// iterate untill diff < epsilon or i_max=7 is reached
// 5 passes converge to <0.25" for the normal operating envelope (alt >= 3deg);
// see testing/check_pointing_inversion.py. Kept a small margin over the bare minimum.
bValid := FALSE;
FOR i:=0 TO 7 BY 1 DO
	d_ha := d_ha_new;
	d_dec := d_dec_new;
	fbpointing(
		HourAngle := LMOD(HourAngle-d_ha,360),
		Declination:= Declination-d_dec,
		Latitude:= Latitude,
		HourAngle_correction => d_ha_new,
		Declination_correction => d_dec_new
	);
	IF ABS(d_ha - d_ha_new) <= epsilon/3600.0 AND ABS(d_dec - d_dec_new) <= epsilon/3600.0 THEN
		bValid := TRUE;
		EXIT;
	END_IF
END_FOR;
// below alt~2-3deg the map is chaotic and never settles within epsilon (see script above);
// do not hand back whatever the last unconverged pass produced
IF bValid THEN
	HourAngle_correction := d_ha_new;
	Declination_correction := d_dec_new;
ELSE
	HourAngle_correction := 0.0;
	Declination_correction := 0.0;
END_IF

END_FUNCTION_BLOCK

// ---- POUs/FB_HomeDropReason.TcPOU
// Why a pending home was dropped after 2 min (#108): the text for the home end state and the WARN. Pure logic,
// tested offline in IAG50cmTests (#120). Order matters: not ready wins over a stop that did not finish.
FUNCTION_BLOCK FB_HomeDropReason
VAR_INPUT
	bReady			: BOOL;		// telescope ready
	bStopPending	: BOOL;		// TCS_command is stop, or the telescope is not at rest
END_VAR
VAR_OUTPUT
	sEnd			: STRING(40);
	sWhy			: STRING(160);
END_VAR

IF NOT bReady THEN
	sEnd := 'cancelled: telescope not ready';
	sWhy := 'the telescope was not ready for 2 min. Power on, then send the home again.';
ELSIF bStopPending THEN
	sEnd := 'cancelled: stop did not finish';
	sWhy := 'the stop before the home did not finish within 2 min. Send the stop, then the home again.';
ELSE
	sEnd := 'cancelled: axes busy';
	sWhy := 'the axes were busy for 2 min. Send the home again.';
END_IF

END_FUNCTION_BLOCK

// ---- POUs/FB_SweepStop.TcPOU
// A stop in the calibration sweep (#113): the axes stay enabled and uncalibrated, the sweep is aborted by the stop. Once the
// stop has settled (for 3 scans) and no homing is running any more, the uncalibrated axes are switched off for one scan, so
// the telescope ends like a stop in the covers phase (READY_STATE -2, no error) and the next power-on starts the sweep
// again. Calibrated axes stay enabled. Pure logic, tested offline in IAG50cmTests.
// #197: ArmAll() is the same for a park without a completed power-on (the axes are on, but the telescope can never be
// ready): every axis is switched off once at rest, calibrated or not, and the axes-off park then parks in place.
FUNCTION_BLOCK FB_SweepStop
VAR_INPUT
	bSettled		: BOOL;		// FB_TelescopeControl.bSettled: at rest and no stop transaction running
	bHaCalibrated	: BOOL;
	bDecCalibrated	: BOOL;
	bHaHoming		: BOOL;		// FB_LatchHome.Busy
	bDecHoming		: BOOL;
	bOtherBusy		: BOOL;		// #197: the focus is moving; waited for in the all-axes mode only
END_VAR
VAR_OUTPUT
	bDisableHa		: BOOL;		// one scan
	bDisableDec		: BOOL;
END_VAR
VAR
	bPending		: BOOL;
	bAll			: BOOL;		// #197: switch every axis off, not only the uncalibrated ones
	nSettledScans	: UINT;
END_VAR
VAR CONSTANT
	nConfirmScans	: UINT := 3;
END_VAR

bDisableHa := FALSE;
bDisableDec := FALSE;
IF bPending THEN
	IF bSettled AND NOT bHaHoming AND NOT bDecHoming AND NOT (bAll AND bOtherBusy) THEN
		IF nSettledScans < nConfirmScans THEN
			nSettledScans := nSettledScans + 1;
		END_IF
	ELSE
		nSettledScans := 0;
	END_IF
	IF nSettledScans >= nConfirmScans THEN
		bDisableHa := bAll OR NOT bHaCalibrated;
		bDisableDec := bAll OR NOT bDecCalibrated;
		bPending := FALSE;
		bAll := FALSE;
	END_IF
END_IF

// A stop arrived in the calibration sweep (power-on stage 40 or later).
METHOD Arm
IF NOT (bPending AND bAll) THEN	// a pending ArmAll() is not narrowed
	bPending := TRUE;
	nSettledScans := 0;
END_IF
END_METHOD

// A park without a completed power-on (#197): switch every axis off once at rest. Idempotent: it may be called every scan.
METHOD ArmAll
IF NOT (bPending AND bAll) THEN
	bPending := TRUE;
	bAll := TRUE;
	nSettledScans := 0;
END_IF
END_METHOD

// Error, reset or a new power-on: nothing to switch off any more.
METHOD Cancel
bPending := FALSE;
bAll := FALSE;
nSettledScans := 0;
END_METHOD

END_FUNCTION_BLOCK

// ---- POUs/Functions/F_HourAngleOffsetOnAxis.TcPOU
// Hour-angle-axis correction (degrees) for a cross-declination offset on the sky (fHourAngleOffset, degrees) at
// declination fDeclination (degrees): fHourAngleOffset / COS(fDeclination). Near the pole 1/COS grows without bound
// and is a division by zero at +-90 deg, so COS is floored at COS(89.5 deg) (factor 115 at most) and the result is
// limited to +-10 deg, the bound BROTLib puts on the offset command (BROTLib#27, same as MONETcommon's
// F_AzimuthOffsetOnAxis near the zenith). Below |dec| = 89.5 deg the result is unchanged.
FUNCTION F_HourAngleOffsetOnAxis : LREAL
VAR_INPUT
	fHourAngleOffset	: LREAL;	// cross-declination offset on the sky, degrees
	fDeclination		: LREAL;	// declination, degrees
END_VAR
VAR CONSTANT
	D2R				: LREAL := 0.017453292519943295;
	MIN_COS			: LREAL := 0.008726535498373935;	// COS(89.5 deg)
	MAX_AXIS_OFFSET	: LREAL := 10.0;					// degrees
END_VAR

F_HourAngleOffsetOnAxis := LIMIT(-MAX_AXIS_OFFSET, fHourAngleOffset / MAX(COS(fDeclination * D2R), MIN_COS), MAX_AXIS_OFFSET);

END_FUNCTION

// ---- POUs/DomeControl/FB_DomeControl.TcPOU
FUNCTION_BLOCK FB_DomeControl IMPLEMENTS I_Dome
VAR_INPUT
	ipTelescope: I_RaDecTelescope;
END_VAR
VAR
	ipState		: I_DomeState := fbDomeIdleState;
	bOpen		: BOOL;
	bClose		: BOOL;
	bReset		: BOOL;
	bHome		: BOOL;
	bTrack		: BOOL;
	bPark		: BOOL;
	bStop		: BOOL;
	bStopDone	: BOOL;
	
	fDomeAziGoInput			: LREAL := 180.0;
	fDomeAziGo				: LREAL := 180.0;
	fDomeAziCurrent			: LREAL := 0.0;
	eDomeRotationState		: E_DomeRotationState;
	eDomeRotationStateOld	: E_DomeRotationState;
	eDomeShutterState		: E_RoofState;
	eDomeShutterStateOld	: E_RoofState;
	bParked			: BOOL;
	
	bDomeError	: BOOL;
	iDomeErrorID: UINT;
	
	ipStateOld			: I_DomeState := fbDomeIdleState;
	fbDomeCloseingState : FB_DomeClosingState(THIS);
	fbDomeErrorState	: FB_DomeErrorState(THIS);
	fbDomeHomeingState	: FB_DomeHomingState(THIS);
	fbDomeIdleState		: FB_DomeIdleState(THIS);
	fbDomeOpeningState	: FB_DomeOpeningState(THIS);
	fbDomeMovingState	: FB_DomeMovingState(THIS);
	fbDomeParkingState	: FB_DomeParkingState(THIS);
	fbDomeStoppingState	: FB_DomeStoppingState(THIS);
	

	rtrigOpen		: R_TRIG;
	rtrigClose		: R_TRIG;
	rtrigReset		: R_TRIG;
	rtrigHome		: R_TRIG;
	rtrigPark		: R_TRIG;
	rtrigStop		: R_TRIG;
	
	fbComm			: I_Comm;
	tonComm 		: TON := (PT:=T#5S);
	
	fbDomeParkedEvent:	FB_EventLog;
	fbDomeStopEvent:	FB_EventLog;
	fbDomeErrorEvent: FB_EventLog;
	
	sSendstring	: STRING;
	Stage		: UINT:= 0;
	Timer		: TON := (PT:=T#30S);
	fbSend		: SendString;
	bSendBusy	: BOOL;
	eSendErrorID: ComError_t;

	fbReceive		: ReceiveString;
	sReceivedString	: STRING;
	sLastReceivedString: STRING;
	bStringReceived	: BOOL;
	bReceiveBusy	: BOOL;
	bReceiveError	: BOOL;
	eReceiveErrorID	: ComError_t;
	bReceiveTimeout	: BOOL;
END_VAR
VAR CONSTANT
	nCapabilities : INT := 2; 	//OPEN TSI : TELESCOPE.CONFIG.CAPABILITIES
END_VAR

// account for off center mount
IF fDomeAziGoInput >= 0.0 AND fDomeAziGoInput < 115.0 THEN
	fDomeAziGo := fDomeAziGoInput - 5.0;
ELSIF fDomeAziGoInput >= 225.0 AND fDomeAziGoInput < 360.0 THEN
	fDomeAziGo := fDomeAziGoInput + 5.0;
ELSE
	fDomeAziGo := fDomeAziGoInput;
END_IF

//	Receive string data:
fbReceive(
	Prefix:='',
	Suffix:= '',
	Timeout:= T#1S,
	ReceivedString:= sReceivedString,
	RXbuffer:= RxBufferDome,
	StringReceived=> bStringReceived,
	Busy=> bReceiveBusy,
	Error=> ,
	RxTimeout=> bReceiveTimeout );
// Check Errors
IF fbSend.Error <> COMERROR_NOERROR THEN
	eSendErrorID := fbSend.Error;
	bDomeError := TRUE;
END_IF
IF fbReceive.Error <> COMERROR_NOERROR THEN
	eReceiveErrorID := fbReceive.Error;
	bDomeError := TRUE;
END_IF

IF bDomeError THEN
	THIS^.ipState.FoundError();
END_IF

rtrigOpen(CLK := bOpen);
rtrigClose(CLK := bClose);
rtrigReset(CLK := bReset);
rtrigHome(CLK := bHome);
rtrigPark(CLK := bPark);
rtrigStop(CLK := bStop);

// #96: a stop wins over every other request of the same scan, which are dropped with it
IF (rtrigStop.Q) THEN
	bStop := FALSE;
	bOpen := FALSE;
	bClose := FALSE;
	bHome := FALSE;
	bPark := FALSE;
	bTrack := FALSE;
	ipState.StopCommand();
END_IF

IF (rtrigReset.Q) THEN
	bReset := FALSE;
	ipState.ResetCommand();
END_IF

IF (rtrigClose.Q) THEN
	bClose := FALSE;
	ipState.CloseCommand();
END_IF

IF (rtrigOpen.Q) THEN
	bOpen := FALSE;
	ipState.OpenCommand();
END_IF

IF (rtrigHome.Q) THEN
	bHome := FALSE;
	ipState.HomeCommand();
END_IF

IF (rtrigPark.Q) THEN
	bPark := FALSE;
	bTrack := FALSE;
	ipState.ParkCommand();
END_IF

// #83: requests are one-shot, like the covers (#66). They are consumed in this scan whether they produced an edge or
// not: a caller repeating a request every scan gave a single edge and then left the flag TRUE, so no later request of
// that kind had an edge until a PLC restart.
bOpen := FALSE;
bClose := FALSE;
bReset := FALSE;
bHome := FALSE;
bPark := FALSE;
bStop := FALSE;

bStopDone := FALSE;
ipState.RunState();

IF eDomeRotationState = E_DomeRotationState.parked AND eDomeShutterState = E_RoofState.closed THEN
	bParked := TRUE;
ELSE
	bParked := FALSE;
END_IF
// send telemetry
tonComm(IN:=TRUE);
IF tonComm.Q THEN // publish new payload every 5 seconds
	tonComm(IN:=FALSE);
	THIS^._SendTelemetry();	
END_IF


fbDomeParkedEvent(
	Trigger := bParked,
	Level := ADSLOG_MSGTYPE_HINT,
	OnMessage := 'Dome is in parking position and closed.',
	comm:= fbComm);
fbDomeStopEvent(
	Trigger := bStopDone,
	Level := ADSLOG_MSGTYPE_HINT,
	OnMessage := 'Dome stopped: rotation holds the current azimuth, a shutter movement is not stopped.',
	comm:= fbComm);
fbDomeErrorEvent(
	Trigger := bDomeError,
	Level := ADSLOG_MSGTYPE_ERROR,
	FormatString := 'Dome Error %s',
	OnMessage := 'found.',
	OffMessage := 'resolved.',
	comm:= fbComm);
// Buffer
ipStateOld := ipState;
eDomeRotationStateOld := eDomeRotationState;
eDomeShutterStateOld := eDomeShutterState;

PROPERTY _DomeRotationState : E_DomeRotationState
GET
_DomeRotationState := eDomeRotationState;
END_GET
SET
eDomeRotationState := _DomeRotationState;
END_SET
END_PROPERTY

PROPERTY _DomeShutterState : E_RoofState
GET
_DomeShutterState := eDomeShutterState;
END_GET
SET
eDomeShutterState := _DomeShutterState;
END_SET
END_PROPERTY

PROPERTY  _Error : BOOL
GET
_Error := bDomeError;
END_GET
SET
bDomeError := _Error;
END_SET
END_PROPERTY

PROPERTY _StopDone : BOOL
GET
_StopDone := bStopDone;
END_GET
SET
bStopDone := _StopDone;
END_SET
END_PROPERTY

PROPERTY _HasReceivedString : Bool
GET
_HasReceivedString := bStringReceived;
END_GET
SET
END_SET
END_PROPERTY

PROPERTY _Parked : BOOL
GET
_Parked := bParked;
END_GET
SET
bParked := _Parked;
END_SET
END_PROPERTY

PROPERTY _Position : LREAL
GET
_Position := fDomeAziGo;
END_GET
SET
fDomeAziCurrent := _Position;
END_SET
END_PROPERTY

PROPERTY _ReceivedString : STRING
GET
_ReceivedString := sReceivedString;
END_GET
SET
END_SET
END_PROPERTY

METHOD _SendTelemetry : BOOL
VAR_INPUT
END_VAR
IF eDomeShutterState = E_RoofState.opened THEN
	fbComm.PublishLREAL('telescope', 'dome', 'AUXILIARY.DOME.REALPOS', 1.0);
ELSIF eDomeShutterState = E_RoofState.closing OR eDomeShutterState = E_RoofState.opening OR eDomeShutterState = E_RoofState.unknown THEN
	fbComm.PublishLREAL('telescope', 'dome', 'AUXILIARY.DOME.REALPOS', 0.5);
ELSIF eDomeShutterState = E_RoofState.closed THEN
	fbComm.PublishLREAL('telescope', 'dome', 'AUXILIARY.DOME.REALPOS', 0.0);
ELSE
	fbComm.PublishLREAL('telescope', 'dome', 'AUXILIARY.DOME.REALPOS', -1.0);
END_IF

IF ipState.StateID = 'Opening State' THEN
	fbComm.PublishLREAL('telescope', 'dome', 'AUXILIARY.DOME.TARGETPOS', 1.0);
ELSE
	fbComm.PublishLREAL('telescope', 'dome', 'AUXILIARY.DOME.TARGETPOS', 0.0);
END_IF

IF bDomeError THEN
	fbComm.PublishINT('telescope', 'dome', 'AUXILIARY.DOME.ERROR_STATE', 1);
	fbComm.PublishLREAL('telescope', 'dome', 'AUXILIARY.DOME.READY_STATE', -1.0);
ELSE
	fbComm.PublishINT('telescope', 'dome', 'AUXILIARY.DOME.ERROR_STATE', 0);
	IF bParked THEN
		fbComm.PublishLREAL('telescope', 'dome', 'AUXILIARY.DOME.READY_STATE', 0.0);
	ELSIF bTrack THEN
		fbComm.PublishLREAL('telescope', 'dome', 'AUXILIARY.DOME.READY_STATE', 8.0);
	ELSE
		fbComm.PublishLREAL('telescope', 'dome', 'AUXILIARY.DOME.READY_STATE', 1.0);
	END_IF
END_IF

IF eDomeRotationState = E_DomeRotationState.slewing OR eDomeRotationState = E_DomeRotationState.unknown THEN
	fbComm.PublishLREAL('telescope', 'dome', 'AUXILIARY.DOME.MOTION_STATE', 1.0);
ELSE
	fbComm.PublishLREAL('telescope', 'dome', 'AUXILIARY.DOME.MOTION_STATE', 0.0);
END_IF
fbComm.PublishLREAL('telescope', 'dome', 'AUXILIARY.DOME.AZ', THIS^.Position);
END_METHOD

PROPERTY _Track : BOOL
GET
_Track := bTrack;
END_GET
END_PROPERTY

PROPERTY Capabilities : INT
GET
Capabilities := nCapabilities;
END_GET
END_PROPERTY

METHOD Close : BOOL
VAR_INPUT
END_VAR
bClose:=True;
END_METHOD

PROPERTY Closed : BOOL
GET
END_GET
END_PROPERTY

PROPERTY Error : Bool
GET
Error := bDomeError;
END_GET
END_PROPERTY

PROPERTY ErrorID : UDINT
GET
END_GET
END_PROPERTY

//FB_Init is always available implicitly and it is used primarily for initialization.
//The return value is not evaluated. For a specific influence, you can also declare the
//methods explicitly and provide additional code there with the standard initialization
//code. You can evaluate the return value.
METHOD FB_Init: BOOL
VAR_INPUT
    bInitRetains	: BOOL; // TRUE: the retain variables are initialized (reset warm / reset cold)
    bInCopyCode		: BOOL;  // TRUE: the instance will be copied to the copy code afterward (online change)
	comm			: I_Comm;
END_VAR
THIS^.fbComm 				:= comm;
END_METHOD

METHOD Open : BOOL
VAR_INPUT
END_VAR
bOpen := True;
END_METHOD

PROPERTY Opened : BOOL
GET
END_GET
END_PROPERTY

METHOD Park : BOOL
VAR_INPUT
END_VAR
bPark := TRUE;
END_METHOD

PROPERTY Parked : BOOL
GET
Parked := bParked;
END_GET
END_PROPERTY

PROPERTY Position : LREAL
GET
Position := fDomeAziCurrent;
END_GET
SET
fDomeAziGoInput := Position;
END_SET
END_PROPERTY

METHOD Reset : BOOL
VAR_INPUT
END_VAR
bReset := True;
END_METHOD

PROPERTY RotState : E_DomeRotationState
GET
RotState := eDomeRotationState;
END_GET
END_PROPERTY

METHOD SetState : BOOL
VAR_INPUT
	newState :I_DomeState;
END_VAR
THIS^.ipState := newState;
END_METHOD

{warning 'add property implementation'}
PROPERTY ShutterState : BROTLib.E_RoofState
GET
END_GET
SET
END_SET
END_PROPERTY

PROPERTY Slewing : BOOL
GET
END_GET
END_PROPERTY

METHOD Stop : BOOL
VAR_INPUT
END_VAR
// #96: the dome has no stop command, the state holds the azimuth it reads (FB_DomeStoppingState)
bStop := TRUE;
END_METHOD

METHOD StopTrack : BOOL
VAR_INPUT
END_VAR
bTrack := FALSE;
END_METHOD

METHOD Track : BOOL
VAR_INPUT
END_VAR
bTrack := TRUE;
END_METHOD

PROPERTY Tracking : BOOL
GET
Tracking := bTrack;
END_GET
END_PROPERTY

END_FUNCTION_BLOCK

// ---- POUs/DomeControl/States/FB_DomeClosingState.TcPOU
FUNCTION_BLOCK FB_DomeClosingState EXTENDS  FB_DomeState
VAR
	Stage		: UINT:= 0;
	tonSleep	: TON := (PT:=T#5S);
	tonTimeout	: TON:= (PT:=T#3M); // see Baader Handbook
	// #202: d#closhut is acknowledged (d#gotmess) but the shutter stays open (d#shutope): the command is sent again at
	// most nMaxAttempts times in all, then it is an error. Before, it was sent for ever, because the timeout is stopped
	// at every poll, and nothing was logged.
	nAttempts	: UINT;
	nMaxAttempts: UINT := 3;
END_VAR


METHOD CloseCommand : BOOL
// #202: a new close starts the shutter command again, with a fresh count
LogEvent(sText := 'Dome: close received while closing, the shutter command is started again', sLevel := 'WARNING');
nAttempts := 0;
Stage := 0;
tonSleep(IN:=FALSE);
tonTimeout(IN:=FALSE);
END_METHOD

METHOD FoundError : BOOL
nAttempts := 0;
Stage:= 0;
tonSleep(IN:=FALSE);
tonTimeout(IN:=FALSE);
pDome^._Error := TRUE;
pDome^.SetState(pDome^.fbDomeErrorState);
END_METHOD


METHOD OpenCommand : BOOL
nAttempts := 0;
Stage:= 0;
tonSleep(IN:=FALSE);
tonTimeout(IN:=FALSE);
pDome^.SetState(pDome^.fbDomeOpeningState);
END_METHOD

METHOD RunState : BOOL
VAR_INPUT
END_VAR
CASE Stage OF
	0:
		tonTimeout(IN:=TRUE);
		Stage := 1;
	1:
		pDome^.fbSend(	SendString:= 'd#closhut',
					TXbuffer:= TxBufferDome,
					Busy=>,
					Error=> );
		IF NOT pDome^.fbSend.Busy  THEN
			Stage := 2;
		END_IF
	2:
		IF pDome^.bStringReceived THEN
			IF pDome^._ReceivedString = 'd#comerro' OR pDome^._ReceivedString = 'd#domerro' THEN
				foundError();
			ELSIF pDome^._ReceivedString = 'd#gotmess' THEN
				Stage := 3;
			END_IF
		ELSIF NOT pDome^.fbReceive.Busy THEN
			tonSleep(IN:=TRUE);
			IF tonSleep.Q THEN
				tonSleep(IN:=FALSE);
				Stage := 1;
			END_IF
		END_IF
		tonTimeout(IN:=TRUE);
		IF tonTimeout.Q THEN
			tonTimeout(IN:=FALSE);
			foundError();
		END_IF
	3:
		tonTimeout(IN:=FALSE);
		
		tonSleep(IN:=TRUE);
		IF tonSleep.Q THEN
			tonSleep(IN:=FALSE);
			Stage := 4;
			tonTimeout(IN:=TRUE);
		END_IF
	4:
		pDome^.fbSend(	SendString:= 'd#getshut',
					TXbuffer:= TxBufferDome,
					Busy=>,
					Error=> );
		IF NOT pDome^.fbSend.Busy  THEN
			Stage := 5;
		END_IF
	5: 
		IF pDome^.bStringReceived THEN
			IF pDome^._ReceivedString = 'd#comerro' OR pDome^._ReceivedString = 'd#domerro' THEN
				FoundError();
			ELSIF pDome^._ReceivedString = 'd#shutclo' THEN
				pDome^._DomeShutterState := E_RoofState.closed;
				Stage := 6;
			ELSIF pDome^._ReceivedString = 'd#shutope' THEN
				pDome^._DomeShutterState := E_RoofState.opened;
				nAttempts := nAttempts + 1;
				IF nAttempts >= nMaxAttempts THEN
					LogEvent(sText := 'Dome: the shutter does not close, d#closhut is acknowledged but the shutter stays open', sLevel := 'WARNING');
					FoundError();
				ELSE
					Stage := 0;
				END_IF
			ELSIF pDome^._ReceivedString = 'd#shutrun' THEN
				pDome^._DomeShutterState := E_RoofState.closing;
				Stage := 3;
			END_IF
		ELSIF NOT pDome^.fbReceive.Busy THEN
			// mixed up string? ask again
			tonSleep(IN:=TRUE);
			IF tonSleep.Q THEN
				tonSleep(IN:=FALSE);
				Stage := 4;
			END_IF
		END_IF
		tonTimeout(IN:=TRUE);
		IF tonTimeout.Q THEN
			tonTimeout(IN:=FALSE);
			FoundError();
		END_IF
	
	6:
		tonTimeout(IN:=FALSE);
		SuccessfulFinished();
		
END_CASE
END_METHOD


PROPERTY StateID : STRING
GET
StateID := 'Closing State';
END_GET
END_PROPERTY


METHOD SuccessfulFinished : BOOL
nAttempts := 0;
Stage:= 0;
tonSleep(IN:=FALSE);
tonTimeout(IN:=FALSE);
pDome^.SetState(pDome^.fbDomeIdleState);
END_METHOD

END_FUNCTION_BLOCK

// ---- POUs/DomeControl/States/FB_DomeState.TcPOU
FUNCTION_BLOCK FB_DomeState IMPLEMENTS I_DomeState

VAR
	TxBuffer	: ComBuffer;
	RxBuffer	: ComBuffer;
	pDome : POINTER TO FB_DomeControl;
END_VAR


METHOD CloseCommand : BOOL
LogIgnored(sCommand := 'close', sLevel := 'WARNING');
END_METHOD

METHOD FB_init : BOOL
VAR_INPUT
	bInitRetains : BOOL; // if TRUE, the retain variables are initialized (warm start / cold start)
	bInCopyCode : BOOL;  // if TRUE, the instance afterwards gets moved into the copy code (online change)
	pDome : POINTER TO FB_DomeControl;

END_VAR
THIS^.pDome := pDome;
END_METHOD


METHOD FoundError : BOOL
END_METHOD


METHOD HomeCommand : BOOL
LogIgnored(sCommand := 'home', sLevel := 'INFO');
END_METHOD

// #202: a line to the ADS log and to 50cm/Log (level WARNING or INFO)
METHOD LogEvent : BOOL
VAR_INPUT
	sText		: STRING(255);
	sLevel		: STRING(20) := 'INFO';
END_VAR
IF sLevel = 'WARNING' THEN
	ADSLOGSTR(ADSLOG_MSGTYPE_WARN OR ADSLOG_MSGTYPE_LOG, '%s', sText);
ELSE
	ADSLOGSTR(ADSLOG_MSGTYPE_HINT OR ADSLOG_MSGTYPE_LOG, '%s', sText);
END_IF
IF pDome <> 0 THEN
	IF pDome^.fbComm <> 0 THEN
		pDome^.fbComm.PublishLog(level := sLevel, message := sText);
	END_IF
END_IF
LogEvent := TRUE;
END_METHOD

// #202: a command that the state does not handle is dropped. Before, it was dropped without a trace: four dome_close
// went unnoticed while the dome was stuck in Closing.
METHOD LogIgnored : BOOL
VAR_INPUT
	sCommand	: STRING(20);
	sLevel		: STRING(20) := 'INFO';
END_VAR
LogIgnored := LogEvent(sText := CONCAT(CONCAT(CONCAT('Dome: ', sCommand), ' ignored in '), THIS^.StateID), sLevel := sLevel);
END_METHOD

METHOD MoveCommand : BOOL
END_METHOD


METHOD OpenCommand : BOOL
LogIgnored(sCommand := 'open', sLevel := 'INFO');
END_METHOD


METHOD ParkCommand : BOOL
LogIgnored(sCommand := 'park', sLevel := 'INFO');
END_METHOD


METHOD ResetCommand : BOOL
LogIgnored(sCommand := 'reset', sLevel := 'INFO');
END_METHOD

METHOD RunState : BOOL
VAR_INPUT
END_VAR
END_METHOD


PROPERTY StateID : STRING
GET
END_GET
END_PROPERTY


METHOD StopCommand : BOOL
LogIgnored(sCommand := 'stop', sLevel := 'INFO');
END_METHOD


METHOD SuccessfulFinished : BOOL
END_METHOD


METHOD TrackCommand : BOOL
END_METHOD

END_FUNCTION_BLOCK

// ---- POUs/DomeControl/States/FB_DomeErrorState.TcPOU
FUNCTION_BLOCK FB_DomeErrorState EXTENDS  FB_DomeState
VAR
END_VAR


METHOD CloseCommand : BOOL
// #202: a close is accepted in every state, it is the way to shut the roof
// the error is cleared like a reset does it: the shutter command must not wait for a dome_reset
ResetCommand();
pDome^.SetState(pDome^.fbDomeCloseingState);
END_METHOD


METHOD ResetCommand : BOOL
VAR
	fbClearTx			: ClearComBuffer;
	fbClearRx			: ClearComBuffer;
END_VAR
fbClearTx(Buffer:=TxBuffer);
fbClearRx(Buffer:=TxBuffer);

pDome^._Error := FALSE;
pDome^.SetState(pDome^.fbDomeIdleState);
END_METHOD


PROPERTY StateID : STRING
GET
StateID := 'Error State';
END_GET
END_PROPERTY

END_FUNCTION_BLOCK

// ---- POUs/DomeControl/States/FB_DomeHomingState.TcPOU
FUNCTION_BLOCK FB_DomeHomingState EXTENDS  FB_DomeState
VAR
END_VAR


METHOD CloseCommand : BOOL
// #202: a close is accepted in every state, it is the way to shut the roof
pDome^.SetState(pDome^.fbDomeCloseingState);
END_METHOD


PROPERTY StateID : STRING
GET
StateID := 'Homing State';
END_GET
END_PROPERTY

END_FUNCTION_BLOCK

// ---- POUs/DomeControl/States/FB_DomeIdleState.TcPOU
FUNCTION_BLOCK FB_DomeIdleState EXTENDS  FB_DomeState

VAR
	Stage		: UINT:= 0;
	tonSleep	: TON := (PT:=T#5S);
	tonTimeout	: TON:= (PT:=T#3M); // see Baader Handbook
	tonDelay	: TON:= (PT:=T#20MS);
	
	sSeperator		: STRING := 'd#azi';
	sLeft			: STRING;
	sAzi			: STRING;
	fAzi			: LREAL;
	fAzi_Old		: LREAL;
	// #202: two azimuth readings closer than this (deg) are the same position: the dome reports tenths of a degree
	// and a single step of jitter must not keep the rotation state at slewing (dome_close is refused while slewing)
	fAziTolerance	: LREAL := 0.5;
	bSplitSuccess 	: BOOL;
	
END_VAR


METHOD CloseCommand : BOOL
IF pDome^._DomeRotationState <> E_DomeRotationState.slewing THEN
	Stage:= 0;
	tonSleep(IN:=FALSE);
	tonTimeout(IN:=FALSE);
	tonDelay(IN:=FALSE);
	pDome^.SetState(pDome^.fbDomeCloseingState);
ELSE
	// #202: not silently. The rotation state is slewing as long as two azimuth readings differ.
	LogIgnored(sCommand := 'close (dome rotating)', sLevel := 'WARNING');
END_IF
END_METHOD


METHOD FoundError : BOOL
Stage:= 0;
tonSleep(IN:=FALSE);
tonTimeout(IN:=FALSE);
tonDelay(IN:=FALSE);
pDome^._Error := TRUE;
pDome^.SetState(pDome^.fbDomeErrorState);
END_METHOD

METHOD MoveCommand : BOOL
Stage:= 0;
tonSleep(IN:=FALSE);
tonTimeout(IN:=FALSE);
tonDelay(IN:=FALSE);
pDome^.SetState(pDome^.fbDomeMovingState);
END_METHOD


METHOD OpenCommand : BOOL
Stage:= 0;
tonSleep(IN:=FALSE);
tonTimeout(IN:=FALSE);
tonDelay(IN:=FALSE);
pDome^.SetState(pDome^.fbDomeOpeningState);
END_METHOD


METHOD ParkCommand : BOOL
Stage:= 0;
tonSleep(IN:=FALSE);
tonTimeout(IN:=FALSE);
tonDelay(IN:=FALSE);
pDome^.SetState(pDome^.fbDomeParkingState);
END_METHOD

METHOD RunState : BOOL
VAR_INPUT
END_VAR
// send 'd#getshut' wait for answer
// wait 5 seconds
// send 'd#getazi' wait for answer
CASE Stage OF
	0:
		tonTimeout(IN:=TRUE);
		Stage := 1;
	1:
		pDome^.fbSend(	SendString:= 'd#getshut',
						TXbuffer:= TxBufferDome,
						Busy=>,
						Error=> );
		IF NOT pDome^.fbSend.Busy  THEN
			Stage := 2;
		END_IF
	2: 
		IF pDome^.bStringReceived THEN
			IF pDome^._ReceivedString = 'd#comerro' OR pDome^._ReceivedString = 'd#domerro' THEN
				FoundError();
			ELSIF pDome^._ReceivedString = 'd#shutclo' THEN
				pDome^._DomeShutterState := E_RoofState.closed;
				Stage := 3;
			ELSIF pDome^._ReceivedString = 'd#shutope' THEN
				pDome^._DomeShutterState := E_RoofState.opened;
				Stage := 3;
			ELSIF pDome^._ReceivedString = 'd#shutrun' THEN
				pDome^._DomeShutterState := E_RoofState.unknown;
				Stage := 3;
			END_IF
		ELSIF NOT pDome^.fbReceive.Busy THEN
			tonSleep(IN:=TRUE);
			IF tonSleep.Q THEN
				tonSleep(IN:=FALSE);
				Stage := 1;
			END_IF
		END_IF
		tonTimeout(IN:=TRUE);
		IF tonTimeout.Q THEN
			tonTimeout(IN:=FALSE);
			FoundError();
		END_IF
	3:
		tonTimeout(IN:=FALSE);
		tonSleep(IN:=TRUE);
		IF tonSleep.Q THEN
			tonSleep(IN:=FALSE);
			Stage := 4;
			tonTimeout(IN:=TRUE);
		END_IF
	4:
		pDome^.fbSend(	SendString:= 'd#getazim',
						TXbuffer:= TxBufferDome,
						Busy=>,
						Error=> );
		IF NOT pDome^.fbSend.Busy  THEN
			Stage := 5;
		END_IF
	5: 
		IF pDome^._HasReceivedString THEN
			IF pDome^._ReceivedString = 'd#comerro' OR pDome^._ReceivedString = 'd#domerro' THEN
				FoundError();
			ELSE
				bSplitSuccess := FindAndSplit(
									pSeparator := ADR(sSeperator),
									pSrcString := ADR(pDome^.sReceivedString),
									pLeftString:= ADR(sLeft),
									nLeftSize	:= 1,
									pRightString := ADR(sAzi),
									nRightSize := 5,
									bSearchFromRight:= FALSE);
									
				IF bSplitSuccess AND ( STRING_TO_LREAL(sAzi) <> 0 OR sAzi = '0000') THEN
					// (STRING_TO_LREAL(sAzi) <> 0 OR sAzi := '0000') -> either sAzi actual 0 OR STRING_TO_LREAL error
					fAzi := STRING_TO_LREAL(sAzi)/10.0;
					//Baader measures azimuth as West of South, so we need to convert it. This works both ways.
					IF fAzi  >= 180.0 THEN
						pDome^._Position := fAzi - 180.0;
					ELSE
						pDome^._Position := fAzi + 180.0;
					END_IF
					IF ABS(fAzi - fAzi_Old) < fAziTolerance THEN
						IF ABS(pDome^.Position - 180.0) < 5.0 THEN
							pDome^._DomeRotationState := E_DomeRotationState.parked;
						ELSE
							pDome^._DomeRotationState := E_DomeRotationState.idle;
						END_IF
					ELSE
						pDome^._DomeRotationState := E_DomeRotationState.slewing;
					END_IF
					fAzi_Old := fAzi;
					Stage := 6;
				END_IF
			END_IF
		ELSIF NOT pDome^.fbReceive.Busy THEN
			tonSleep(IN:=TRUE);
			IF tonSleep.Q THEN
				tonSleep(IN:=FALSE);
				Stage := 4;
			END_IF
		END_IF
		tonTimeout(IN:=TRUE);
		IF tonTimeout.Q THEN
			tonTimeout(IN:=FALSE);
			FoundError();
		END_IF
	6:
		tonTimeout(IN:=FALSE);
		IF ABS( pDome^.Position - pDome^._Position) > 10.0 AND pDome^._Track THEN
			MoveCommand();
		ELSE
			Stage:= 7;
		END_IF
	7:
		tonSleep(IN:=TRUE);
		IF tonSleep.Q THEN
			tonSleep(IN:=FALSE);
			Stage := 0;
		END_IF		
END_CASE
END_METHOD


METHOD StopCommand : BOOL
Stage:= 0;
tonSleep(IN:=FALSE);
tonTimeout(IN:=FALSE);
tonDelay(IN:=FALSE);
pDome^.SetState(pDome^.fbDomeStoppingState);
END_METHOD


PROPERTY StateID : STRING
GET
StateID := 'Idle State';
END_GET
END_PROPERTY

END_FUNCTION_BLOCK

// ---- POUs/DomeControl/States/FB_DomeOpeningState.TcPOU
FUNCTION_BLOCK FB_DomeOpeningState EXTENDS  FB_DomeState

VAR
	Stage		: UINT:= 0;
	tonSleep	: TON := (PT:=T#2S);
	tonTimeout	: TON:= (PT:=T#3M); // see Baader Handbook
	// #202: d#opeshut acknowledged but the shutter reports closed: at most nMaxAttempts sends in all, then an error
	nAttempts	: UINT;
	nMaxAttempts: UINT := 3;
END_VAR


METHOD CloseCommand : BOOL
nAttempts := 0;
Stage := 0;
tonSleep(IN:=FALSE);
tonTimeout(IN:=FALSE);
pDome^.SetState(pDome^.fbDomeCloseingState);
END_METHOD


METHOD FoundError : BOOL
nAttempts := 0;
Stage := 0;
tonSleep(IN:=FALSE);
tonTimeout(IN:=FALSE);
pDome^._Error := TRUE;
pDome^.SetState(pDome^.fbDomeErrorState);
END_METHOD

METHOD RunState : BOOL
VAR_INPUT
END_VAR
CASE Stage OF
	0:
		tonTimeout(IN:=TRUE);
		Stage := 1;
	1:
		pDome^.fbSend(	SendString:= 'd#opeshut',
					TXbuffer:= TxBufferDome,
					Busy=>,
					Error=> );
		IF NOT pDome^.fbSend.Busy  THEN
			Stage := 2;
		END_IF
	2:
		IF pDome^.bStringReceived THEN
			IF pDome^._ReceivedString = 'd#comerro' OR pDome^._ReceivedString = 'd#domerro' THEN
				FoundError();
			ELSIF pDome^._ReceivedString = 'd#gotmess' THEN
				Stage := 3;
			END_IF
		ELSIF NOT pDome^.fbReceive.Busy THEN
			tonSleep(IN:=TRUE);
			IF tonSleep.Q THEN
				tonSleep(IN:=FALSE);
				Stage := 1;
			END_IF
		END_IF
		tonTimeout(IN:=TRUE);
		IF tonTimeout.Q THEN
			tonTimeout(IN:=FALSE);
			FoundError();
		END_IF
	3:
		tonTimeout(IN:=FALSE);
		tonSleep(IN:=TRUE);
		IF tonSleep.Q THEN
			tonSleep(IN:=FALSE);
			Stage := 4;
			tonTimeout(IN:=TRUE);
		END_IF
	4:
		pDome^.fbSend(	SendString:= 'd#getshut',
					TXbuffer:= TxBufferDome,
					Busy=>,
					Error=> );
		IF NOT pDome^.fbSend.Busy  THEN
			Stage := 5;
		END_IF
	5: 
		IF pDome^.bStringReceived THEN
			IF pDome^._ReceivedString = 'd#comerro' OR pDome^._ReceivedString = 'd#domerro' THEN
				FoundError();
			ELSIF pDome^._ReceivedString = 'd#shutclo' THEN
				pDome^._DomeShutterState := E_RoofState.closed;
				tonTimeout(IN:=FALSE);
				nAttempts := nAttempts + 1;
				IF nAttempts >= nMaxAttempts THEN
					LogEvent(sText := 'Dome: the shutter does not open, d#opeshut is acknowledged but the shutter stays closed', sLevel := 'WARNING');
					FoundError();
				ELSE
					Stage := 0; // restart
				END_IF
			ELSIF pDome^._ReceivedString = 'd#shutope' THEN
				pDome^._DomeShutterState := E_RoofState.opened;
				Stage := 6;
			ELSIF pDome^._ReceivedString = 'd#shutrun' THEN
				pDome^._DomeShutterState := E_RoofState.opening;
				Stage := 3; // wait longer
			END_IF
		ELSIF NOT pDome^.fbReceive.Busy THEN
			tonSleep(IN:=TRUE);
			IF tonSleep.Q THEN
				tonSleep(IN:=FALSE);
				Stage := 4;
			END_IF
		END_IF
		
		tonTimeout(IN:=TRUE);
		IF tonTimeout.Q THEN
			tonTimeout(IN:=FALSE);
			FoundError();
		END_IF
	
	6:
		tonTimeout(IN:=FALSE);
		SuccessfulFinished();
END_CASE
END_METHOD


PROPERTY StateID : STRING
GET
StateID := 'Opening State';
END_GET
END_PROPERTY


METHOD SuccessfulFinished : BOOL
nAttempts := 0;
Stage := 0;
tonSleep(IN:=FALSE);
tonTimeout(IN:=FALSE);
pDome^.SetState(pDome^.fbDomeIdleState);
END_METHOD

END_FUNCTION_BLOCK

// ---- POUs/DomeControl/States/FB_DomeMovingState.TcPOU
FUNCTION_BLOCK FB_DomeMovingState EXTENDS  FB_DomeState

VAR
	Stage		: UINT:= 0;
	tonSleep	: TON := (PT:=T#5S);
	tonTimeout	: TON:= (PT:=T#3M); // see Baader Handbook
	tonDelay	: TON:= (PT:=T#20MS);
	tonMoveDelay: TON:= (PT:=T#10M); // only move the Dome every PT minutes
	
	sSeperator		: STRING := 'd#azi';
	sSend			: STRING := 'd#azi';
	sLeft			: STRING;
	sAzi			: STRING;
	fAzi		: LREAL;
	fAzi_Old		: LREAL;
	bSplitSuccess 	: BOOL;
END_VAR


METHOD CloseCommand : BOOL
// #202: a close is accepted in every state, it is the way to shut the roof
Stage := 0;
tonSleep(IN:=FALSE);
tonTimeout(IN:=FALSE);
tonDelay(IN:=FALSE);
pDome^.SetState(pDome^.fbDomeCloseingState);
END_METHOD


METHOD FoundError : BOOL
Stage:= 0;
tonSleep(IN:=FALSE);
tonTimeout(IN:=FALSE);
tonDelay(IN:=FALSE);
pDome^._Error := TRUE;
pDome^.SetState(pDome^.fbDomeErrorState);
END_METHOD


METHOD ParkCommand : BOOL
Stage:= 0;
tonSleep(IN:=FALSE);
tonTimeout(IN:=FALSE);
tonDelay(IN:=FALSE);
pDome^.SetState(pDome^.fbDomeParkingState);
END_METHOD

METHOD RunState : BOOL
VAR_INPUT
END_VAR
CASE Stage OF
	0:
		tonTimeout(IN:=TRUE);
		Stage:=1;
	1:
		//Baader measures azimuth as West of South, so we need to convert it. This works both ways.
		
		IF pDome^._Position  >= 180.0 THEN
			fAzi := pDome^._Position - 180.0;
		ELSE
			fAzi := pDome^._Position + 180.0;
		END_IF
		IF LREAL_TO_INT(fAzi*10) < 10 THEN
			sSend := CONCAT('d#azi000',  INT_TO_STRING(LREAL_TO_INT(fAzi*10)));
		ELSIF LREAL_TO_INT(fAzi*10) < 100 THEN
			sSend := CONCAT('d#azi00',  INT_TO_STRING(LREAL_TO_INT(fAzi*10)));
		ELSIF LREAL_TO_INT(fAzi*10) < 1000 THEN
			sSend := CONCAT('d#azi0',  INT_TO_STRING(LREAL_TO_INT(fAzi*10)));
		ELSE
			sSend := CONCAT('d#azi', INT_TO_STRING(LREAL_TO_INT(fAzi*10)));
		END_IF
		pDome^.fbSend(	SendString:= sSend,
					TXbuffer:= TxBufferDome,
					Busy=>,
					Error=> );
		IF NOT pDome^.fbSend.Busy  THEN
			Stage := 2;
		END_IF
	2: 
		IF pDome^._HasReceivedString THEN
			pDome^._DomeRotationState := E_DomeRotationState.slewing;
			IF pDome^._ReceivedString = 'd#comerro' OR pDome^._ReceivedString = 'd#domerro' THEN
				FoundError();
			ELSIF  pDome^._ReceivedString = 'd#gotmess' THEN
				Stage := 3;
			END_IF
		ELSIF NOT pDome^.fbReceive.Busy THEN
			tonSleep(IN:=TRUE);
			IF tonSleep.Q THEN
				tonSleep(IN:=FALSE);
				Stage := 1;
			END_IF
		END_IF
		tonTimeout(IN:=TRUE);
		IF tonTimeout.Q THEN
			tonTimeout(IN:=FALSE);
			FoundError();
		END_IF
	3:
		SuccessfulFinished();
END_CASE
END_METHOD


PROPERTY StateID : STRING
GET
StateID := 'Moving State';
END_GET
END_PROPERTY


METHOD StopCommand : BOOL
Stage:= 0;
tonSleep(IN:=FALSE);
tonTimeout(IN:=FALSE);
tonDelay(IN:=FALSE);
pDome^.SetState(pDome^.fbDomeStoppingState);
END_METHOD

METHOD SuccessfulFinished : BOOL
Stage := 0;
tonSleep(IN:=FALSE);
tonTimeout(IN:=FALSE);
pDome^.SetState(pDome^.fbDomeIdleState);
END_METHOD

END_FUNCTION_BLOCK

// ---- POUs/DomeControl/States/FB_DomeParkingState.TcPOU
FUNCTION_BLOCK FB_DomeParkingState EXTENDS FB_DomeState

VAR
	Stage		: UINT:= 0;
	tonTimeout	: TON:= (PT:=T#3M); // see Baader Handbook
	tonSleep	: TON := (PT:=T#2S);
	tonDelay	: TON:= (PT:=T#20MS);
	
	sSeperator		: STRING := 'd#azi';
	sLeft			: STRING;
	sAzi			: STRING;
	fAzi			: LREAL;
	fAzi_Old		: LREAL;
	bSplitSuccess 	: BOOL;
END_VAR


METHOD CloseCommand : BOOL
Stage := 0;
tonSleep(IN:=FALSE);
tonTimeout(IN:=FALSE);
tonDelay(IN:=FALSE);
pDome^.SetState(pDome^.fbDomeCloseingState);
END_METHOD


METHOD FoundError : BOOL
Stage:= 0;
tonSleep(IN:=FALSE);
tonTimeout(IN:=FALSE);
tonDelay(IN:=FALSE);
pDome^._Error := TRUE;
pDome^.SetState(pDome^.fbDomeErrorState);
END_METHOD

METHOD OpenCommand : BOOL
Stage:= 0;
tonSleep(IN:=FALSE);
tonTimeout(IN:=FALSE);
tonDelay(IN:=FALSE);
pDome^.SetState(pDome^.fbDomeOpeningState);
END_METHOD

METHOD RunState : BOOL
VAR_INPUT
END_VAR
CASE Stage OF
	0:
		tonTimeout(IN:=TRUE);
		IF NOT pDome^.fbReceive.Busy AND NOT pDome^.fbSend.Busy THEN
			Stage := 1;
		END_IF
	1:
		pDome^.fbSend(	SendString:= 'd#azi0000',
					TXbuffer:= TxBufferDome,
					Busy=>,
					Error=> );
		IF NOT pDome^.fbSend.Busy  THEN
			Stage := 2;
		END_IF
	2:
		IF pDome^._HasReceivedString THEN
			IF pDome^._ReceivedString = 'd#comerro' OR pDome^._ReceivedString = 'd#domerro' THEN
				FoundError();
			ELSIF pDome^._ReceivedString = 'd#gotmess' THEN
				Stage := 3;
			END_IF
		ELSIF NOT pDome^.fbReceive.Busy THEN
			tonSleep(IN:=TRUE);
			IF tonSleep.Q THEN
				tonSleep(IN:=FALSE);
				Stage := 1;
			END_IF
		END_IF
		tonTimeout(IN:=TRUE);
		IF tonTimeout.Q THEN
			tonTimeout(IN:=FALSE);
			FoundError();
		END_IF
	3:
		tonTimeout(IN:=FALSE);
		tonSleep(IN:=TRUE);
		IF tonSleep.Q THEN
			tonSleep(IN:=FALSE);
			Stage := 4;
			tonTimeout(IN:=TRUE);
		END_IF
	4:
		pDome^.fbSend(	SendString:= 'd#getazim',
					TXbuffer:= TxBufferDome,
					Busy=>,
					Error=> );
		IF NOT pDome^.fbSend.Busy  THEN
			Stage := 5;
		END_IF
	5: 
		IF pDome^._HasReceivedString THEN
			IF pDome^._ReceivedString = 'd#comerro' OR pDome^._ReceivedString = 'd#domerro' THEN
				FoundError();
			ELSE
				bSplitSuccess := FindAndSplit(
									pSeparator := ADR(sSeperator),
									pSrcString := ADR(pDome^.sReceivedString),
									pLeftString:= ADR(sLeft),
									nLeftSize	:= 1,
									pRightString := ADR(sAzi),
									nRightSize := 5,
									bSearchFromRight:= FALSE);
				IF bSplitSuccess AND ( STRING_TO_LREAL(sAzi) <> 0 OR sAzi = '0000' ) THEN
					// (STRING_TO_LREAL(sAzi) <> 0 OR sAzi := '0000') -> either sAzi actual 0 OR STRING_TO_LREAL error
					fAzi := STRING_TO_LREAL(sAzi)/10.0;
					//Baader measures azimuth as West of South, so we need to convert it. This works both ways.
					IF fAzi  >= 180.0 THEN
						pDome^._Position := fAzi - 180.0;
					ELSE
						pDome^._Position := fAzi + 180.0;
					END_IF
					IF fAzi = fAzi_Old THEN
						IF ABS(pDome^.Position - 180.0) < 5.0 THEN
							pDome^._DomeRotationState := E_DomeRotationState.parked;
							Stage := 6;
						ELSE
							pDome^._DomeRotationState := E_DomeRotationState.idle;
							// stopped but not parked? try again
							Stage := 0;
						END_IF
					ELSE
						pDome^._DomeRotationState := E_DomeRotationState.slewing;
						// carry on
						Stage := 3;
					END_IF
					fAzi_Old := fAzi;
				END_IF
			END_IF
		ELSIF NOT pDome^.fbReceive.Busy THEN
			tonSleep(IN:=TRUE);
			IF tonSleep.Q THEN
				tonSleep(IN:=FALSE);
				Stage := 4;
			END_IF
		END_IF
		tonTimeout(IN:=TRUE);
		IF tonTimeout.Q THEN
			tonTimeout(IN:=FALSE);
			FoundError();
		END_IF
	6:
		tonTimeout(IN:=FALSE);
		SuccessfulFinished();
		
END_CASE
END_METHOD

PROPERTY StateID : STRING
GET
StateID := 'Parking State';
END_GET
END_PROPERTY


METHOD StopCommand : BOOL
Stage:= 0;
tonSleep(IN:=FALSE);
tonTimeout(IN:=FALSE);
tonDelay(IN:=FALSE);
pDome^.SetState(pDome^.fbDomeStoppingState);
END_METHOD


METHOD SuccessfulFinished : BOOL
Stage:= 0;
tonSleep(IN:=FALSE);
tonTimeout(IN:=FALSE);
tonDelay(IN:=FALSE);
pDome^.SetState(pDome^.fbDomeIdleState);
END_METHOD

END_FUNCTION_BLOCK

// ---- POUs/DomeControl/States/FB_DomeStoppingState.TcPOU
FUNCTION_BLOCK FB_DomeStoppingState EXTENDS FB_DomeState
// #96: the Baader dome has no stop command. The azimuth target is replaced at once by a new one (manual, page 5), so
// a stop reads the azimuth the dome has now and sends it back as the new target. The azimuth is sent exactly as
// the dome reported it (tenths of a degree, 0000 south): no conversion, no off-centre correction. A shutter
// movement cannot be stopped this way and goes on.
VAR
	Stage		: UINT:= 0;
	tonTimeout	: TON:= (PT:=T#30S);
	tonSleep	: TON := (PT:=T#1S);

	sSeperator		: STRING := 'd#azi';
	sLeft			: STRING;
	sAzi			: STRING;
	bSplitSuccess 	: BOOL;
END_VAR


METHOD CloseCommand : BOOL
// #202: a close is accepted in every state, it is the way to shut the roof
Stage := 0;
tonSleep(IN:=FALSE);
tonTimeout(IN:=FALSE);
pDome^.SetState(pDome^.fbDomeCloseingState);
END_METHOD


METHOD FoundError : BOOL
Stage:= 0;
tonSleep(IN:=FALSE);
tonTimeout(IN:=FALSE);
pDome^._Error := TRUE;
pDome^.SetState(pDome^.fbDomeErrorState);
END_METHOD

METHOD RunState : BOOL
VAR_INPUT
END_VAR
// the stop does not wait for the old move or its 3 min timeout: it is a short transaction of its own
tonTimeout(IN:=TRUE);
IF tonTimeout.Q THEN
	FoundError();
	RETURN;
END_IF

CASE Stage OF
	0:
		// the state that was left may have a request or a reply on the line
		IF NOT pDome^.fbReceive.Busy AND NOT pDome^.fbSend.Busy THEN
			Stage := 1;
		END_IF
	1:
		pDome^.fbSend(	SendString:= 'd#getazim',
					TXbuffer:= TxBufferDome,
					Busy=>,
					Error=> );
		IF NOT pDome^.fbSend.Busy  THEN
			Stage := 2;
		END_IF
	2:
		IF pDome^._HasReceivedString THEN
			IF pDome^._ReceivedString = 'd#comerro' OR pDome^._ReceivedString = 'd#domerro' THEN
				FoundError();
			ELSE
				// a late reply of the cancelled move (d#gotmess) does not split and is waited out
				bSplitSuccess := FindAndSplit(
									pSeparator := ADR(sSeperator),
									pSrcString := ADR(pDome^.sReceivedString),
									pLeftString:= ADR(sLeft),
									nLeftSize	:= 1,
									pRightString := ADR(sAzi),
									nRightSize := 5,
									bSearchFromRight:= FALSE);
				IF bSplitSuccess AND LEN(sAzi) = 4 AND ( STRING_TO_LREAL(sAzi) <> 0 OR sAzi = '0000' ) THEN
					Stage := 3;
				END_IF
			END_IF
		ELSIF NOT pDome^.fbReceive.Busy THEN
			tonSleep(IN:=TRUE);
			IF tonSleep.Q THEN
				tonSleep(IN:=FALSE);
				Stage := 1;
			END_IF
		END_IF
	3:
		pDome^.fbSend(	SendString:= CONCAT('d#azi', sAzi),
					TXbuffer:= TxBufferDome,
					Busy=>,
					Error=> );
		IF NOT pDome^.fbSend.Busy  THEN
			Stage := 4;
		END_IF
	4:
		IF pDome^._HasReceivedString THEN
			IF pDome^._ReceivedString = 'd#comerro' OR pDome^._ReceivedString = 'd#domerro' THEN
				FoundError();
			ELSIF pDome^._ReceivedString = 'd#gotmess' THEN
				SuccessfulFinished();
			END_IF
		ELSIF NOT pDome^.fbReceive.Busy THEN
			tonSleep(IN:=TRUE);
			IF tonSleep.Q THEN
				tonSleep(IN:=FALSE);
				Stage := 3;
			END_IF
		END_IF
END_CASE
END_METHOD


PROPERTY StateID : STRING
GET
StateID := 'Stopping State';
END_GET
END_PROPERTY

METHOD SuccessfulFinished : BOOL
Stage := 0;
tonSleep(IN:=FALSE);
tonTimeout(IN:=FALSE);
pDome^._DomeRotationState := E_DomeRotationState.idle;
pDome^._StopDone := TRUE;
pDome^.SetState(pDome^.fbDomeIdleState);
END_METHOD

END_FUNCTION_BLOCK

// ---- POUs/PendantControl/FB_PendantControl.TcPOU
FUNCTION_BLOCK FB_PendantControl
VAR_INPUT
	ipTelescope	: I_RaDecTelescope;
	ipFocus		: I_Focus;
END_VAR
VAR_OUTPUT
END_VAR
VAR
	fbComm			: I_Comm;
	tonComm 		: TON := (PT:=T#5S);
	(*  State Definitions *)
	ipState			: I_PendantState := fbPendantPreInitState;
	ipStateOld		: I_PendantState := fbPendantPreInitState;
	
	fbPendantPreInitState	: FB_PendantPreInitState(THIS);
	fbPendantIdleState 		: FB_PendantIdleState(THIS);
	fbPendantInitState 		: FB_PendantInitState(THIS);
	fbPendantSetHAState		: FB_PendantSetHAState(THIS);
	fbPendantSetDECState	: FB_PendantSetDECState(THIS);
	fbPendantSetFocusState	: FB_PendantSetFocusState(THIS);
	fbPendantErrorState		: FB_PendantErrorState(THIS);
	
	bReady			: BOOL;
	bError			: BOOL;
	bReset			: BOOL;
	nErrorID		: UINT;
	
	(* Set Logic:
		bFastMove:	TRUE (move big step)
					FALSE (move small step)
		bMovePositive:	TRUE +
						FALSE -*)
	bFastMove		: BOOL;
	bMovePositive	: BOOL;
	
	rtrigReset		: R_TRIG;
	rtrigError		: R_TRIG;
	
	(*SEND*)
	fbSendString	: SendString;
	fbSendHex		: SendData;
	eSendErrorID	: ComError_t;
	
	
	(* RECEIVE*)
	fbReceive		: ReceiveString;
	rtrigReceive	: R_TRIG;
	sReceivedString	: STRING;
	sLastReceivedString: STRING;
	bStringReceived	: BOOL;
	bReceiveBusy	: BOOL;
	bReceiveError	: BOOL;
	eReceiveErrorID	: ComError_t;
	bReceiveTimeout	: BOOL;
END_VAR

//	Receive string data:	
fbReceive(
	Prefix:='',
	Suffix:= '',
	Timeout:= T#1MS,
	ReceivedString:= sReceivedString,
	RXbuffer:= RxBufferPendant,
	StringReceived=> bStringReceived,
	Busy=> bReceiveBusy,
	Error=> ,
	RxTimeout=> bReceiveTimeout );

(*Send / Receive Errors? *)
IF fbReceive.Error <> COMERROR_NOERROR THEN
	bError:=TRUE;
	nErrorID		:= fbReceive.Error;
	eReceiveErrorID := fbReceive.Error;
END_IF
IF fbSendString.Error <> COMERROR_NOERROR THEN
	bError:=TRUE;
	nErrorID	:= fbSendString.Error;
	eSendErrorID := fbSendString.Error;
ELSIF fbSendHex.Error <> COMERROR_NOERROR THEN
	bError:=TRUE;
	nErrorID := fbSendHex.Error;
	eSendErrorID := fbSendHex.Error;
END_IF

(* Triggers*)
rtrigReceive(CLK:=bStringReceived);
rtrigReset(CLK:=bReset);
rtrigError(CLK:=bError);

IF rtrigError.Q THEN
	bFastMove := FALSE;
	ipState.FoundError();
ELSIF rtrigReset.Q THEN
	ipState.ResetCommand();
	bReset:=FALSE;
ELSIF rtrigReceive.Q AND NOT bError THEN
	(* INIT *)
	IF sReceivedString = '#' THEN
		ipState.InitCommand();
		
	(* HA *)
	ELSIF sReceivedString = 'û' AND bReady THEN
		(* -, slow*)
		bFastMove := FALSE;
		bMovePositive := FALSE;
		ipState.HaCommand();
	ELSIF sReceivedString = '{' AND bReady THEN
		(* -, fast*)
		bFastMove := TRUE;
		bMovePositive := FALSE;
		ipState.HaCommand();
	ELSIF sReceivedString = 'ý' AND bReady THEN
		(* +, slow*)
		bFastMove := FALSE;
		bMovePositive := TRUE;
		ipState.HaCommand();
	ELSIF sReceivedString = '}' AND bReady THEN
		(* +, fast*)
		bFastMove := TRUE;
		bMovePositive := TRUE;
		ipState.HaCommand();
	
	(* DEC *)
	ELSIF sReceivedString = 'ï' AND bReady THEN
		(* -, slow*)
		bFastMove := FALSE;
		bMovePositive := FALSE;
		ipState.DecCommand();
	ELSIF sReceivedString = 'o' AND bReady THEN
		(* -, fast*)
		bFastMove := TRUE;
		bMovePositive := FALSE;
		ipState.DecCommand();
	ELSIF sReceivedString = '÷' AND bReady THEN
		(* +, slow*)
		bFastMove := FALSE;
		bMovePositive := TRUE;
		ipState.DecCommand();
	ELSIF sReceivedString = 'w' AND bReady THEN
		(* +, fast*)
		bFastMove := TRUE;
		bMovePositive := TRUE;
		ipState.DecCommand();
	
	(* Focus *)
	ELSIF sReceivedString = '¿' AND bReady THEN
		(* -, slow*)
		bFastMove := FALSE;
		bMovePositive := FALSE;
		ipState.FocusCommand();
	ELSIF sReceivedString = '?' AND bReady THEN
		(* -, fast*)
		bFastMove := TRUE;
		bMovePositive := FALSE;
		ipState.FocusCommand();
	ELSIF sReceivedString = 'ß' AND bReady THEN
		(* +, slow*)
		bFastMove := FALSE;
		bMovePositive := TRUE;
		ipState.FocusCommand();
	ELSIF sReceivedString = '_' AND bReady THEN
		(* +, fast*)
		bFastMove := TRUE;
		bMovePositive := TRUE;
		ipState.FocusCommand();
	ELSE
		bFastMove := FALSE;
		ipState.ToIdle();
	END_IF
	
END_IF

ipState.RunState();

PROPERTY _Error : BOOL
GET
_Error := bError;
END_GET
SET
bError:=_Error;
END_SET
END_PROPERTY

PROPERTY _FastMove : BOOL
GET
_FastMove := THIS^.bFastMove;
END_GET
END_PROPERTY

PROPERTY _MovePositive : BOOL
GET
_MovePositive := THIS^.bMovePositive;
END_GET
END_PROPERTY

PROPERTY _Ready : BOOL
GET
_Ready := bReady;
END_GET
SET
bReady := _Ready;
END_SET
END_PROPERTY

PROPERTY Error : BOOL
GET
Error := bError;
END_GET
END_PROPERTY

PROPERTY ErrorID : UINT
GET
ErrorID := nErrorID;
END_GET
END_PROPERTY

//FB_Init is always available implicitly and it is used primarily for initialization.
//The return value is not evaluated. For a specific influence, you can also declare the
//methods explicitly and provide additional code there with the standard initialization
//code. You can evaluate the return value.
METHOD FB_Init: BOOL
VAR_INPUT
    bInitRetains	: BOOL; // TRUE: the retain variables are initialized (reset warm / reset cold)
    bInCopyCode		: BOOL;  // TRUE: the instance will be copied to the copy code afterward (online change)
	comm			: I_Comm;
END_VAR
THIS^.fbComm 				:= comm;
END_METHOD

PROPERTY Reset : BOOL
SET
bReset := Reset;
END_SET
END_PROPERTY

METHOD SetState : BOOL
VAR_INPUT
	newState :I_PendantState;
END_VAR
THIS^.ipState := newState;
END_METHOD

END_FUNCTION_BLOCK

// ---- POUs/PendantControl/States/FB_PendantPreInitState.TcPOU
FUNCTION_BLOCK FB_PendantPreInitState EXTENDS FB_PendantState
VAR_INPUT
END_VAR
VAR_OUTPUT
END_VAR
VAR
END_VAR

METHOD FoundError : BOOL
pPendant^.SetState(pPendant^.fbPendantErrorState);
END_METHOD

METHOD InitCommand : BOOL
pPendant^.SetState(pPendant^.fbPendantInitState);
END_METHOD

PROPERTY StateID : STRING
GET
StateID := 'Pre Init State';
END_GET
END_PROPERTY

END_FUNCTION_BLOCK

// ---- POUs/PendantControl/States/FB_PendantState.TcPOU
FUNCTION_BLOCK FB_PendantState IMPLEMENTS I_PendantState
VAR
	TxBuffer	: ComBuffer;
	RxBuffer	: ComBuffer;
	pPendant : POINTER TO FB_PendantControl;
END_VAR

{warning 'add method implementation '}
METHOD DecCommand : BOOL
END_METHOD

METHOD FB_init : BOOL
VAR_INPUT
	bInitRetains : BOOL; // if TRUE, the retain variables are initialized (warm start / cold start)
	bInCopyCode : BOOL;  // if TRUE, the instance afterwards gets moved into the copy code (online change)
	pPendant : POINTER TO FB_PendantControl;

END_VAR
THIS^.pPendant := pPendant;
END_METHOD

{warning 'add method implementation '}
METHOD FocusCommand : BOOL
END_METHOD

{warning 'add method implementation '}
METHOD FoundError : BOOL
END_METHOD

{warning 'add method implementation '}
METHOD HaCommand : BOOL
END_METHOD

{warning 'add method implementation '}
METHOD InitCommand : BOOL
END_METHOD

{warning 'add method implementation '}
METHOD ResetCommand : BOOL
END_METHOD

{warning 'add method implementation '}
METHOD RunState : BOOL
END_METHOD

{warning 'add property implementation'}
PROPERTY StateID : STRING
GET
END_GET
END_PROPERTY

{warning 'add method implementation '}
METHOD Timeout : BOOL
END_METHOD

{warning 'add method implementation '}
METHOD ToIdle : BOOL
END_METHOD

END_FUNCTION_BLOCK

// ---- POUs/PendantControl/States/FB_PendantIdleState.TcPOU
FUNCTION_BLOCK FB_PendantIdleState EXTENDS FB_PendantState
VAR_INPUT
END_VAR
VAR_OUTPUT
END_VAR
VAR
	Stage			: UINT:= 0;
	bBlockChange	: BOOL := FALSE;
	tonSleep		: TON := (PT:=T#10S);
	
	fHaOffset		: LREAL;
	sHaOffset		: STRING;
	sHaOffsetLeft	: STRING;
	sHaOffsetRight	: STRING;
	nHaOffsetLength	: INT;
	nHaOffsetRightLength :INT;
	
	fDecOffset		: LREAL;
	sDecOffset		: STRING;
	sDecOffsetLeft	: STRING;
	sDecOffsetRight	: STRING;
	nDecOffsetLength: INT;
	nDecOffsetRightLength :INT;
	
	fFocusPosition	: LREAL;
	sFocusPosition	: STRING;
	nFocusRightLength :INT;
	
	
	//Hex stuff
	aTxHexData		: ARRAY[0..2] OF BYTE;
	tonDelay		: TON:= (PT:=T#20MS);
END_VAR

METHOD DecCommand : BOOL
IF NOT bBlockChange THEN
	Stage := 0;
	tonDelay(IN:=FALSE);
	tonSleep(IN:=FALSE);
	pPendant^.SetState(pPendant^.fbPendantSetDecState);
END_IF
END_METHOD

METHOD FocusCommand : BOOL
IF NOT bBlockChange THEN
	Stage := 0;
	tonDelay(IN:=FALSE);
	tonSleep(IN:=FALSE);
	pPendant^.SetState(pPendant^.fbPendantSetFocusState);
END_IF
END_METHOD

METHOD FoundError : BOOL
Stage := 0;
tonDelay(IN:=FALSE);
tonSleep(IN:=FALSE);
bBlockChange:= FALSE;
pPendant^.SetState(pPendant^.fbPendantErrorState);
END_METHOD

METHOD HaCommand : BOOL
IF NOT bBlockChange THEN
	Stage := 0;
	tonDelay(IN:=FALSE);
	tonSleep(IN:=FALSE);
	pPendant^.SetState(pPendant^.fbPendantSetHaState);
END_IF
END_METHOD

METHOD InitCommand : BOOL
IF NOT bBlockChange THEN
	Stage := 0;
	tonDelay(IN:=FALSE);
	tonSleep(IN:=FALSE);
	pPendant^.SetState(pPendant^.fbPendantInitState);
END_IF
END_METHOD

METHOD RunState : BOOL
(*---- IDLE----
	Show:	Ha :**** "
			Dec:**** "
	Sleep
	
	Show:	Fokus (1-17mm)
			******** mm
	Sleep
	-> repeat
*)
CASE Stage OF
	0:
		tonSleep(IN:=TRUE);
		IF tonSleep.Q THEN
			tonSleep(IN:=FALSE);
			Stage:=Stage +1;
		END_IF
	1:
		// Block State Change while full text is send -> to not run into issues with commands
		// Does not include Error State
		bBlockChange := TRUE;
		IF NOT pPendant^.fbSendHex.Busy OR pPendant^.fbSendString.Busy THEN
			Stage := Stage +1;
		END_IF
	2: 
		// send sequence for two line text. For first line: fe, 01, 00, 0c, first 8 char, second 8 char
		HEXSTR_TO_DATA('fe', ADR(aTxHexData), SIZEOF(aTxHexData));
		pPendant^.fbSendHex(
				pSendData:= ADR(aTxHexData),
				Length	:= 1,
				TXbuffer:= TxBufferPendant,
				Busy=>,
				Error=> );
		IF NOT pPendant^.fbSendHex.Busy THEN
			Stage := Stage +1;
		END_IF
	3: 
		HEXSTR_TO_DATA('01', ADR(aTxHexData), SIZEOF(aTxHexData));
		pPendant^.fbSendHex(
				pSendData:= ADR(aTxHexData),
				Length	:= 1,
				TXbuffer:= TxBufferPendant,
				Busy=>,
				Error=> );
		IF NOT pPendant^.fbSendHex.Busy THEN
			Stage := Stage +1;
		END_IF
	4: 
		HEXSTR_TO_DATA('00', ADR(aTxHexData), SIZEOF(aTxHexData));
		pPendant^.fbSendHex(
				pSendData:= ADR(aTxHexData),
				Length	:= 1,
				TXbuffer:= TxBufferPendant,
				Busy=>,
				Error=> );
		IF NOT pPendant^.fbSendHex.Busy THEN
			Stage := Stage +1;
		END_IF
	5:	
		HEXSTR_TO_DATA('0c', ADR(aTxHexData), SIZEOF(aTxHexData));
		pPendant^.fbSendHex(
				pSendData:= ADR(aTxHexData),
				Length	:= 1,
				TXbuffer:= TxBufferPendant,
				Busy=>,
				Error=> );
		IF NOT pPendant^.fbSendHex.Busy THEN
			Stage := Stage +1;
		END_IF
	6:
		// Get Offset
		fHaOffset := F_RoundLREAL(pPendant^.ipTelescope.HourAngleOffset*3600,0);
		sHaOffset := INT_TO_STRING(LREAL_TO_INT(fHaOffset));
		nHaOffsetLength := LEN(sHaOffset);
		// needs to be devided into 8 + rest characters
		IF nHaOffsetLength < 4 THEN
			sHaOffsetLeft := sHaOffset;
			IF nHaOffsetLength < 3 THEN
				sHaOffsetLeft := CONCAT(sHaOffsetLeft, '"');
				sHaOffsetRight:='       .';
			ELSE
				sHaOffsetRight:='"       ';
			END_IF
		ELSE
			sHaOffsetLeft := Left(sHaOffset,3);
			sHaOffsetRight := CONCAT(CONCAT(Right(sHaOffset, nHaOffsetLength-3), '"'),'        ');
		END_IF
		IF fHaOffset >= 0 THEN
			sHaOffsetLeft := CONCAT('+', sHaOffsetLeft);
		END_IF
		// send first 8 characters
		pPendant^.fbSendString(SendString:= CONCAT('HA :',sHaOffsetLeft ),
					TXbuffer:= TxBufferPendant,
					Busy=>,
					Error=> );
		IF NOT pPendant^.fbSendString.Busy  THEN
			Stage := Stage +1;
		END_IF
	7: 
		tonDelay(IN:=TRUE);
		IF tonDelay.Q THEN
			tonDelay(IN:=FALSE);
			Stage:=Stage +1;
		END_IF
	8:
		// send second 8 characters
		pPendant^.fbSendString(SendString:= MID(sHaOffsetRight,8,1),
					TXbuffer:= TxBufferPendant,
					Busy=>,
					Error=> );
		IF NOT pPendant^.fbSendString.Busy  THEN
			Stage := Stage +1;
		END_IF
	9: 
		tonDelay(IN:=TRUE);
		IF tonDelay.Q THEN
			tonDelay(IN:=FALSE);
			Stage:=Stage +1;
		END_IF
	10:
		// second line: fe, c0, 00, 0b, first 8 char, second 8 char
		HEXSTR_TO_DATA('fe', ADR(aTxHexData), SIZEOF(aTxHexData));
		pPendant^.fbSendHex(
				pSendData:= ADR(aTxHexData),
				Length	:= 1,
				TXbuffer:= TxBufferPendant,
				Busy=>,
				Error=> );
		IF NOT pPendant^.fbSendHex.Busy THEN
			Stage := Stage +1;
		END_IF
	11: 
		HEXSTR_TO_DATA('c0', ADR(aTxHexData), SIZEOF(aTxHexData));
		pPendant^.fbSendHex(
				pSendData:= ADR(aTxHexData),
				Length	:= 1,
				TXbuffer:= TxBufferPendant,
				Busy=>,
				Error=> );
		IF NOT pPendant^.fbSendHex.Busy THEN
			Stage := Stage +1;
		END_IF
	12: 
		HEXSTR_TO_DATA('00', ADR(aTxHexData), SIZEOF(aTxHexData));
		pPendant^.fbSendHex(
				pSendData:= ADR(aTxHexData),
				Length	:= 1,
				TXbuffer:= TxBufferPendant,
				Busy=>,
				Error=> );
		IF NOT pPendant^.fbSendHex.Busy THEN
			Stage := Stage +1;
		END_IF
	13:	
		HEXSTR_TO_DATA('0b', ADR(aTxHexData), SIZEOF(aTxHexData));
		pPendant^.fbSendHex(
				pSendData:= ADR(aTxHexData),
				Length	:= 1,
				TXbuffer:= TxBufferPendant,
				Busy=>,
				Error=> );
		IF NOT pPendant^.fbSendHex.Busy THEN
			Stage := Stage +1;
		END_IF
	14:
		fDecOffset := F_RoundLREAL(pPendant^.ipTelescope.DeclinationOffset*3600,0);
		sDecOffset := INT_TO_STRING(LREAL_TO_INT(fDecOffset));
		nDecOffsetLength := LEN(sDecOffset);
		IF nDecOffsetLength < 4 THEN
			sDecOffsetLeft := sDecOffset;
			IF nDecOffsetLength < 3 THEN
				sDecOffsetLeft := CONCAT(sDecOffsetLeft, '"');
				sDecOffsetRight:='       .';
			ELSE
				sDecOffsetRight:='"      .';
			END_IF
		ELSE
			sDecOffsetLeft := Left(sDecOffset,3);
			sDecOffsetRight := CONCAT(CONCAT(Right(sDecOffset, nDecOffsetLength-3), '"'),'        ');
		END_IF
		IF fDecOffset >= 0 THEN
			sDecOffsetLeft := CONCAT('+', sDecOffsetLeft);
		END_IF
		
		pPendant^.fbSendString(SendString:= CONCAT('Dec:',sDecOffsetLeft ),
					TXbuffer:= TxBufferPendant,
					Busy=>,
					Error=> );
		IF NOT pPendant^.fbSendString.Busy  THEN
			Stage := Stage +1;
		END_IF
	15: 
		tonDelay(IN:=TRUE);
		IF tonDelay.Q THEN
			tonDelay(IN:=FALSE);
			Stage:=Stage +1;
		END_IF
	16:
		pPendant^.fbSendString(SendString:=MID(sDecOffsetRight,8,1),
					TXbuffer:= TxBufferPendant,
					Busy=>,
					Error=> );
		IF NOT pPendant^.fbSendString.Busy  THEN
			// unblock State change
			bBlockChange := FALSE;
			Stage := Stage +1;
		END_IF
	17:
		// Sleep for some time
		tonSleep(IN:=TRUE);
		IF tonSleep.Q THEN
			tonSleep(IN:=FALSE);
			Stage:=Stage +1;
		END_IF
	18:
		// Block State Change while full text is send -> to not run into issues with commands
		// Does not include Error State
		bBlockChange := TRUE;
		IF NOT pPendant^.fbSendHex.Busy OR pPendant^.fbSendString.Busy THEN
			Stage := Stage +1;
		END_IF
	19: 
		// send sequence for two line text. For first line: fe, 01, 00, 0c, first 8 char, second 8 char
		HEXSTR_TO_DATA('fe', ADR(aTxHexData), SIZEOF(aTxHexData));
		pPendant^.fbSendHex(
				pSendData:= ADR(aTxHexData),
				Length	:= 1,
				TXbuffer:= TxBufferPendant,
				Busy=>,
				Error=> );
		IF NOT pPendant^.fbSendHex.Busy THEN
			Stage := Stage +1;
		END_IF
	20: 
		HEXSTR_TO_DATA('01', ADR(aTxHexData), SIZEOF(aTxHexData));
		pPendant^.fbSendHex(
				pSendData:= ADR(aTxHexData),
				Length	:= 1,
				TXbuffer:= TxBufferPendant,
				Busy=>,
				Error=> );
		IF NOT pPendant^.fbSendHex.Busy THEN
			Stage := Stage +1;
		END_IF
	21: 
		HEXSTR_TO_DATA('00', ADR(aTxHexData), SIZEOF(aTxHexData));
		pPendant^.fbSendHex(
				pSendData:= ADR(aTxHexData),
				Length	:= 1,
				TXbuffer:= TxBufferPendant,
				Busy=>,
				Error=> );
		IF NOT pPendant^.fbSendHex.Busy THEN
			Stage := Stage +1;
		END_IF
	22:	
		HEXSTR_TO_DATA('0c', ADR(aTxHexData), SIZEOF(aTxHexData));
		pPendant^.fbSendHex(
				pSendData:= ADR(aTxHexData),
				Length	:= 1,
				TXbuffer:= TxBufferPendant,
				Busy=>,
				Error=> );
		IF NOT pPendant^.fbSendHex.Busy THEN
			Stage := Stage +1;
		END_IF
	23:
		// send first 8 characters
		pPendant^.fbSendString(SendString:= 'Focus 1-',
					TXbuffer:= TxBufferPendant,
					Busy=>,
					Error=> );
		IF NOT pPendant^.fbSendString.Busy  THEN
			Stage := Stage +1;
		END_IF
	24: 
		tonDelay(IN:=TRUE);
		IF tonDelay.Q THEN
			tonDelay(IN:=FALSE);
			Stage:=Stage +1;
		END_IF
	25:
		// send second characters (8 max)
		pPendant^.fbSendString(SendString:= '17mm    ',
					TXbuffer:= TxBufferPendant,
					Busy=>,
					Error=> );
		IF NOT pPendant^.fbSendString.Busy  THEN
			Stage := Stage +1;
		END_IF
	26: 
		tonDelay(IN:=TRUE);
		IF tonDelay.Q THEN
			tonDelay(IN:=FALSE);
			Stage:=Stage +1;
		END_IF
	27: 
		// second line: fe, c0, 00, 0b, first 8 char, second 8 char
		HEXSTR_TO_DATA('fe', ADR(aTxHexData), SIZEOF(aTxHexData));
		pPendant^.fbSendHex(
				pSendData:= ADR(aTxHexData),
				Length	:= 1,
				TXbuffer:= TxBufferPendant,
				Busy=>,
				Error=> );
		IF NOT pPendant^.fbSendHex.Busy THEN
			Stage := Stage +1;
		END_IF
	28: 
		HEXSTR_TO_DATA('c0', ADR(aTxHexData), SIZEOF(aTxHexData));
		pPendant^.fbSendHex(
				pSendData:= ADR(aTxHexData),
				Length	:= 1,
				TXbuffer:= TxBufferPendant,
				Busy=>,
				Error=> );
		IF NOT pPendant^.fbSendHex.Busy THEN
			Stage := Stage +1;
		END_IF
	29: 
		HEXSTR_TO_DATA('00', ADR(aTxHexData), SIZEOF(aTxHexData));
		pPendant^.fbSendHex(
				pSendData:= ADR(aTxHexData),
				Length	:= 1,
				TXbuffer:= TxBufferPendant,
				Busy=>,
				Error=> );
		IF NOT pPendant^.fbSendHex.Busy THEN
			Stage := Stage +1;
		END_IF
	30:	
		HEXSTR_TO_DATA('0b', ADR(aTxHexData), SIZEOF(aTxHexData));
		pPendant^.fbSendHex(
				pSendData:= ADR(aTxHexData),
				Length	:= 1,
				TXbuffer:= TxBufferPendant,
				Busy=>,
				Error=> );
		IF NOT pPendant^.fbSendHex.Busy THEN
			Stage := Stage +1;
		END_IF
	31:
		// Get Focus Position
		fFocusPosition := F_RoundLREAL(pPendant^.ipFocus.Position,3);
		sFocusPosition := CONCAT(LREAL_TO_STRING(fFocusPosition),'        ');
		// send first 8 characters
		pPendant^.fbSendString(SendString:= MID(sFocusPosition,8,1),
					TXbuffer:= TxBufferPendant,
					Busy=>,
					Error=> );
		IF NOT pPendant^.fbSendString.Busy  THEN
			Stage := Stage +1;
		END_IF
	32: 
		tonDelay(IN:=TRUE);
		IF tonDelay.Q THEN
			tonDelay(IN:=FALSE);
			Stage:=Stage +1;
		END_IF
	33:
		pPendant^.fbSendString(SendString:= 'mm      ',
					TXbuffer:= TxBufferPendant,
					Busy=>,
					Error=> );
		IF NOT pPendant^.fbSendString.Busy  THEN
			// unblock State change
			bBlockChange := FALSE;
			// restart
			Stage := 0;
		END_IF
END_CASE
END_METHOD

PROPERTY StateID : STRING
GET
StateID := 'Idle State';
END_GET
END_PROPERTY

END_FUNCTION_BLOCK

// ---- POUs/PendantControl/States/FB_PendantInitState.TcPOU
FUNCTION_BLOCK FB_PendantInitState EXTENDS FB_PendantState
VAR_INPUT
END_VAR
VAR_OUTPUT
END_VAR
VAR
	Stage		: UINT:= 0;
	
	//Hex stuff
	aTxHexData		: ARRAY[0..2] OF BYTE;
	tonDelay		: TON:= (PT:=T#20MS);

END_VAR

METHOD FoundError : BOOL
Stage := 0;
tonDelay(IN:=FALSE);
pPendant^.SetState(pPendant^.fbPendantErrorState);
END_METHOD

METHOD RunState : BOOL
CASE Stage OF
	0:
		IF NOT pPendant^.fbSendHex.Busy OR pPendant^.fbSendString.Busy THEN
			Stage := Stage +1;
		END_IF
	1:
		HEXSTR_TO_DATA('fd', ADR(aTxHexData), SIZEOF(aTxHexData));
		pPendant^.fbSendHex(
				pSendData:= ADR(aTxHexData),
				Length	:= 1,
				TXbuffer:= TxBufferPendant,
				Busy=>,
				Error=> );
		IF NOT pPendant^.fbSendHex.Busy THEN
			Stage := Stage +1;
		END_IF
	2: 
		
		HEXSTR_TO_DATA('fe', ADR(aTxHexData), SIZEOF(aTxHexData));
		pPendant^.fbSendHex(
				pSendData:= ADR(aTxHexData),
				Length	:= 1,
				TXbuffer:= TxBufferPendant,
				Busy=>,
				Error=> );
		IF NOT pPendant^.fbSendHex.Busy THEN
			Stage := Stage +1;
		END_IF
	3: 
		
		HEXSTR_TO_DATA('01', ADR(aTxHexData), SIZEOF(aTxHexData));
		pPendant^.fbSendHex(
				pSendData:= ADR(aTxHexData),
				Length	:= 1,
				TXbuffer:= TxBufferPendant,
				Busy=>,
				Error=> );
		IF NOT pPendant^.fbSendHex.Busy THEN
			Stage := Stage +1;
		END_IF
	4: 
		
		HEXSTR_TO_DATA('00', ADR(aTxHexData), SIZEOF(aTxHexData));
		pPendant^.fbSendHex(
				pSendData:= ADR(aTxHexData),
				Length	:= 1,
				TXbuffer:= TxBufferPendant,
				Busy=>,
				Error=> );
		IF NOT pPendant^.fbSendHex.Busy THEN
			Stage := Stage +1;
		END_IF
	5:	
		HEXSTR_TO_DATA('0e', ADR(aTxHexData), SIZEOF(aTxHexData));
		pPendant^.fbSendHex(
				pSendData:= ADR(aTxHexData),
				Length	:= 1,
				TXbuffer:= TxBufferPendant,
				Busy=>,
				Error=> );
		IF NOT pPendant^.fbSendHex.Busy THEN
			Stage := Stage +1;
		END_IF
	6:
		pPendant^.fbSendString(SendString:= 'Pendant ',
					TXbuffer:= TxBufferPendant,
					Busy=>,
					Error=> );
		IF NOT pPendant^.fbSendString.Busy  THEN
			Stage := Stage +1;
		END_IF
	7: 
		tonDelay(IN:=TRUE);
		IF tonDelay.Q THEN
			tonDelay(IN:=FALSE);
			Stage:=Stage +1;
		END_IF
	8:
		pPendant^.fbSendString(SendString:= 'on      ',
					TXbuffer:= TxBufferPendant,
					Busy=>,
					Error=> );
		IF NOT pPendant^.fbSendString.Busy  THEN
			Stage := Stage +1;
		END_IF
	9:
		pPendant^._Ready := TRUE;
		THIS^.ToIdle();
END_CASE
END_METHOD

PROPERTY StateID : STRING
GET
StateID := 'Init State';
END_GET
END_PROPERTY

METHOD ToIdle : BOOL
Stage := 0;
pPendant^.SetState(pPendant^.fbPendantIdleState);
END_METHOD

END_FUNCTION_BLOCK

// ---- POUs/PendantControl/States/FB_PendantSetHAState.TcPOU
FUNCTION_BLOCK FB_PendantSetHAState EXTENDS FB_PendantState
VAR_INPUT
END_VAR
VAR_OUTPUT
END_VAR
VAR
		Stage 					: UINT;
	tonCount 				: TON:= (PT:=T#1S);
	fSmallStep				: LREAL := 10;
	fBigStep				: LREAL := 100;
	
	fCurrentHaOffset		: LREAL;
	fSetHaOffset			: LREAL;
	sSetHaOffset			: STRING;
	
	bBlockChange			: BOOL := FALSE;
	bToIdle					: BOOL := FALSE;
	//Hex stuff
	aTxHexData				: ARRAY[0..2] OF BYTE;
	tonDelay				: TON:= (PT:=T#20MS);
END_VAR

METHOD FoundError : BOOL
Stage := 0;
tonDelay(IN:=FALSE);
tonCount(IN:=FALSE);
pPendant^.SetState(pPendant^.fbPendantErrorState);
END_METHOD

METHOD RunState : BOOL
CASE Stage OF
	0:
		fCurrentHaOffset := F_RoundLREAL(pPendant^.ipTelescope.HourAngleOffset*3600,0);
		IF pPendant^._FastMove THEN
			IF pPendant^._MovePositive THEN
				fSetHaOffset := fCurrentHaOffset + fBigStep;
			ELSE
				fSetHaOffset := fCurrentHaOffset - fBigStep;
			END_IF
		ELSE
			IF pPendant^._MovePositive THEN
				fSetHaOffset := fCurrentHaOffset + fSmallStep;
			ELSE
				fSetHaOffset := fCurrentHaOffset - fSmallStep;
			END_IF
		END_IF
		pPendant^.ipTelescope.HourAngleOffset := fSetHaOffset/3600;
		Stage := Stage +1;
	1:
		// Block State Change while full text is send -> to not run into issues with commands
		// Does not include Error State
		bBlockChange := TRUE;
		IF NOT pPendant^.fbSendHex.Busy OR pPendant^.fbSendString.Busy THEN
			Stage := Stage +1;
		END_IF
	2: 
		// send sequence for two line text. For first line: fe, 01, 00, 0c, first 8 char, second 8 char
		HEXSTR_TO_DATA('fe', ADR(aTxHexData), SIZEOF(aTxHexData));
		pPendant^.fbSendHex(
				pSendData:= ADR(aTxHexData),
				Length	:= 1,
				TXbuffer:= TxBufferPendant,
				Busy=>,
				Error=> );
		IF NOT pPendant^.fbSendHex.Busy THEN
			Stage := Stage +1;
		END_IF
	3: 
		HEXSTR_TO_DATA('01', ADR(aTxHexData), SIZEOF(aTxHexData));
		pPendant^.fbSendHex(
				pSendData:= ADR(aTxHexData),
				Length	:= 1,
				TXbuffer:= TxBufferPendant,
				Busy=>,
				Error=> );
		IF NOT pPendant^.fbSendHex.Busy THEN
			Stage := Stage +1;
		END_IF
	4: 
		HEXSTR_TO_DATA('00', ADR(aTxHexData), SIZEOF(aTxHexData));
		pPendant^.fbSendHex(
				pSendData:= ADR(aTxHexData),
				Length	:= 1,
				TXbuffer:= TxBufferPendant,
				Busy=>,
				Error=> );
		IF NOT pPendant^.fbSendHex.Busy THEN
			Stage := Stage +1;
		END_IF
	5:	
		HEXSTR_TO_DATA('0c', ADR(aTxHexData), SIZEOF(aTxHexData));
		pPendant^.fbSendHex(
				pSendData:= ADR(aTxHexData),
				Length	:= 1,
				TXbuffer:= TxBufferPendant,
				Busy=>,
				Error=> );
		IF NOT pPendant^.fbSendHex.Busy THEN
			Stage := Stage +1;
		END_IF
	6:
		// send first 8 characters
		pPendant^.fbSendString(SendString:= 'Ha Offse',
					TXbuffer:= TxBufferPendant,
					Busy=>,
					Error=> );
		IF NOT pPendant^.fbSendString.Busy  THEN
			Stage := Stage +1;
		END_IF
	7: 
		tonDelay(IN:=TRUE);
		IF tonDelay.Q THEN
			tonDelay(IN:=FALSE);
			Stage:=Stage +1;
		END_IF
	8:
		// send second characters (8 max)
		pPendant^.fbSendString(SendString:= 't:      ',
					TXbuffer:= TxBufferPendant,
					Busy=>,
					Error=> );
		IF NOT pPendant^.fbSendString.Busy  THEN
			Stage := Stage +1;
		END_IF
	9: 
		tonDelay(IN:=TRUE);
		IF tonDelay.Q THEN
			tonDelay(IN:=FALSE);
			Stage:=Stage +1;
		END_IF
	10: 
		// second line: fe, c0, 00, 0b, first 8 char, second 8 char
		HEXSTR_TO_DATA('fe', ADR(aTxHexData), SIZEOF(aTxHexData));
		pPendant^.fbSendHex(
				pSendData:= ADR(aTxHexData),
				Length	:= 1,
				TXbuffer:= TxBufferPendant,
				Busy=>,
				Error=> );
		IF NOT pPendant^.fbSendHex.Busy THEN
			Stage := Stage +1;
		END_IF
	11: 
		HEXSTR_TO_DATA('c0', ADR(aTxHexData), SIZEOF(aTxHexData));
		pPendant^.fbSendHex(
				pSendData:= ADR(aTxHexData),
				Length	:= 1,
				TXbuffer:= TxBufferPendant,
				Busy=>,
				Error=> );
		IF NOT pPendant^.fbSendHex.Busy THEN
			Stage := Stage +1;
		END_IF
	12: 
		HEXSTR_TO_DATA('00', ADR(aTxHexData), SIZEOF(aTxHexData));
		pPendant^.fbSendHex(
				pSendData:= ADR(aTxHexData),
				Length	:= 1,
				TXbuffer:= TxBufferPendant,
				Busy=>,
				Error=> );
		IF NOT pPendant^.fbSendHex.Busy THEN
			Stage := Stage +1;
		END_IF
	13:	
		HEXSTR_TO_DATA('0b', ADR(aTxHexData), SIZEOF(aTxHexData));
		pPendant^.fbSendHex(
				pSendData:= ADR(aTxHexData),
				Length	:= 1,
				TXbuffer:= TxBufferPendant,
				Busy=>,
				Error=> );
		IF NOT pPendant^.fbSendHex.Busy THEN
			Stage := Stage +1;
		END_IF
	14:
		IF fSetHaOffset >= 0 THEN
			sSetHaOffset := CONCAT(CONCAT('+',INT_TO_STRING(LREAL_TO_INT(fSetHaOffset))),'        ');
		ELSE
			sSetHaOffset := CONCAT(INT_TO_STRING(LREAL_TO_INT(fSetHaOffset)),'        ');
		END_IF
		
		// send first 8 characters
		pPendant^.fbSendString(SendString:= MID(sSetHaOffset,8,1),
					TXbuffer:= TxBufferPendant,
					Busy=>,
					Error=> );
		IF NOT pPendant^.fbSendString.Busy  THEN
			Stage := Stage +1;
		END_IF
	15: 
		tonDelay(IN:=TRUE);
		IF tonDelay.Q THEN
			tonDelay(IN:=FALSE);
			Stage:=Stage +1;
		END_IF
	16:
		pPendant^.fbSendString(SendString:= '"       ',
					TXbuffer:= TxBufferPendant,
					Busy=>,
					Error=> );
		IF NOT pPendant^.fbSendString.Busy  THEN
			// unblock State change
			bBlockChange := FALSE;
			Stage := Stage +1;
		END_IF
	17:
		tonCount(IN:=TRUE);
		IF tonCount.Q THEN
			tonCount(IN:=FALSE);
			//restart
			Stage:=0;
		END_IF
END_CASE

IF bToIdle THEN
	THIS^.ToIdle();
END_IF
END_METHOD

PROPERTY StateID : STRING
GET
StateID := 'Set Ha Offset State';
END_GET
END_PROPERTY

METHOD ToIdle : BOOL
IF NOT bBlockChange THEN
	Stage := 0;
	tonDelay(IN:=FALSE);
	tonCount(IN:=FALSE);
	bToIdle := FALSE;
	pPendant^.SetState(pPendant^.fbPendantIdleState);
ELSE
	bToIdle := TRUE;
END_IF
END_METHOD

END_FUNCTION_BLOCK

// ---- POUs/PendantControl/States/FB_PendantSetDECState.TcPOU
FUNCTION_BLOCK FB_PendantSetDecState EXTENDS FB_PendantState
VAR_INPUT
END_VAR
VAR_OUTPUT
END_VAR
VAR
	Stage 					: UINT;
	tonCount 				: TON:= (PT:=T#1S);
	fSmallStep				: LREAL := 10;
	fBigStep				: LREAL := 100;
	
	fCurrentDecOffset		: LREAL;
	fSetDecOffset			: LREAL;
	sSetDecOffset			: STRING;
	
	bBlockChange			: BOOL := FALSE;
	bToIdle					: BOOL := FALSE;
	//Hex stuff
	aTxHexData				: ARRAY[0..2] OF BYTE;
	tonDelay				: TON:= (PT:=T#20MS);
END_VAR

METHOD FoundError : BOOL
Stage := 0;
tonDelay(IN:=FALSE);
tonCount(IN:=FALSE);
pPendant^.SetState(pPendant^.fbPendantErrorState);
END_METHOD

METHOD RunState : BOOL
CASE Stage OF
	0:
		fCurrentDecOffset := F_RoundLREAL(pPendant^.ipTelescope.DeclinationOffset*3600,0);
		IF pPendant^._FastMove THEN
			IF pPendant^._MovePositive THEN
				fSetDecOffset := fCurrentDecOffset + fBigStep;
			ELSE
				fSetDecOffset := fCurrentDecOffset - fBigStep;
			END_IF
		ELSE
			IF pPendant^._MovePositive THEN
				fSetDecOffset := fCurrentDecOffset + fSmallStep;
			ELSE
				fSetDecOffset := fCurrentDecOffset - fSmallStep;
			END_IF
		END_IF
		pPendant^.ipTelescope.DeclinationOffset := fSetDecOffset/3600;
		Stage := Stage +1;
	1:
		// Block State Change while full text is send -> to not run into issues with commands
		// Does not include Error State
		bBlockChange := TRUE;
		IF NOT pPendant^.fbSendHex.Busy OR pPendant^.fbSendString.Busy THEN
			Stage := Stage +1;
		END_IF
	2: 
		// send sequence for two line text. For first line: fe, 01, 00, 0c, first 8 char, second 8 char
		HEXSTR_TO_DATA('fe', ADR(aTxHexData), SIZEOF(aTxHexData));
		pPendant^.fbSendHex(
				pSendData:= ADR(aTxHexData),
				Length	:= 1,
				TXbuffer:= TxBufferPendant,
				Busy=>,
				Error=> );
		IF NOT pPendant^.fbSendHex.Busy THEN
			Stage := Stage +1;
		END_IF
	3: 
		HEXSTR_TO_DATA('01', ADR(aTxHexData), SIZEOF(aTxHexData));
		pPendant^.fbSendHex(
				pSendData:= ADR(aTxHexData),
				Length	:= 1,
				TXbuffer:= TxBufferPendant,
				Busy=>,
				Error=> );
		IF NOT pPendant^.fbSendHex.Busy THEN
			Stage := Stage +1;
		END_IF
	4: 
		HEXSTR_TO_DATA('00', ADR(aTxHexData), SIZEOF(aTxHexData));
		pPendant^.fbSendHex(
				pSendData:= ADR(aTxHexData),
				Length	:= 1,
				TXbuffer:= TxBufferPendant,
				Busy=>,
				Error=> );
		IF NOT pPendant^.fbSendHex.Busy THEN
			Stage := Stage +1;
		END_IF
	5:	
		HEXSTR_TO_DATA('0c', ADR(aTxHexData), SIZEOF(aTxHexData));
		pPendant^.fbSendHex(
				pSendData:= ADR(aTxHexData),
				Length	:= 1,
				TXbuffer:= TxBufferPendant,
				Busy=>,
				Error=> );
		IF NOT pPendant^.fbSendHex.Busy THEN
			Stage := Stage +1;
		END_IF
	6:
		// send first 8 characters
		pPendant^.fbSendString(SendString:= 'Dec Offs',
					TXbuffer:= TxBufferPendant,
					Busy=>,
					Error=> );
		IF NOT pPendant^.fbSendString.Busy  THEN
			Stage := Stage +1;
		END_IF
	7: 
		tonDelay(IN:=TRUE);
		IF tonDelay.Q THEN
			tonDelay(IN:=FALSE);
			Stage:=Stage +1;
		END_IF
	8:
		// send second characters (8 max)
		pPendant^.fbSendString(SendString:= 'et:     ',
					TXbuffer:= TxBufferPendant,
					Busy=>,
					Error=> );
		IF NOT pPendant^.fbSendString.Busy  THEN
			Stage := Stage +1;
		END_IF
	9: 
		tonDelay(IN:=TRUE);
		IF tonDelay.Q THEN
			tonDelay(IN:=FALSE);
			Stage:=Stage +1;
		END_IF
	10: 
		// second line: fe, c0, 00, 0b, first 8 char, second 8 char
		HEXSTR_TO_DATA('fe', ADR(aTxHexData), SIZEOF(aTxHexData));
		pPendant^.fbSendHex(
				pSendData:= ADR(aTxHexData),
				Length	:= 1,
				TXbuffer:= TxBufferPendant,
				Busy=>,
				Error=> );
		IF NOT pPendant^.fbSendHex.Busy THEN
			Stage := Stage +1;
		END_IF
	11: 
		HEXSTR_TO_DATA('c0', ADR(aTxHexData), SIZEOF(aTxHexData));
		pPendant^.fbSendHex(
				pSendData:= ADR(aTxHexData),
				Length	:= 1,
				TXbuffer:= TxBufferPendant,
				Busy=>,
				Error=> );
		IF NOT pPendant^.fbSendHex.Busy THEN
			Stage := Stage +1;
		END_IF
	12: 
		HEXSTR_TO_DATA('00', ADR(aTxHexData), SIZEOF(aTxHexData));
		pPendant^.fbSendHex(
				pSendData:= ADR(aTxHexData),
				Length	:= 1,
				TXbuffer:= TxBufferPendant,
				Busy=>,
				Error=> );
		IF NOT pPendant^.fbSendHex.Busy THEN
			Stage := Stage +1;
		END_IF
	13:	
		HEXSTR_TO_DATA('0b', ADR(aTxHexData), SIZEOF(aTxHexData));
		pPendant^.fbSendHex(
				pSendData:= ADR(aTxHexData),
				Length	:= 1,
				TXbuffer:= TxBufferPendant,
				Busy=>,
				Error=> );
		IF NOT pPendant^.fbSendHex.Busy THEN
			Stage := Stage +1;
		END_IF
	14:
		IF fSetDecOffset >= 0 THEN
			sSetDecOffset := CONCAT(CONCAT('+',INT_TO_STRING(LREAL_TO_INT(fSetDecOffset))),'        ');
		ELSE
			sSetDecOffset := CONCAT(INT_TO_STRING(LREAL_TO_INT(fSetDecOffset)),'        ');
		END_IF
		
		// send first 8 characters
		pPendant^.fbSendString(SendString:= MID(sSetDecOffset,8,1),
					TXbuffer:= TxBufferPendant,
					Busy=>,
					Error=> );
		IF NOT pPendant^.fbSendString.Busy  THEN
			Stage := Stage +1;
		END_IF
	15: 
		tonDelay(IN:=TRUE);
		IF tonDelay.Q THEN
			tonDelay(IN:=FALSE);
			Stage:=Stage +1;
		END_IF
	16:
		pPendant^.fbSendString(SendString:= '"       ',
					TXbuffer:= TxBufferPendant,
					Busy=>,
					Error=> );
		IF NOT pPendant^.fbSendString.Busy  THEN
			// unblock State change
			bBlockChange := FALSE;
			Stage := Stage +1;
		END_IF
	17:
		tonCount(IN:=TRUE);
		IF tonCount.Q THEN
			tonCount(IN:=FALSE);
			//restart
			Stage:=0;
		END_IF
END_CASE

IF bToIdle THEN
	THIS^.ToIdle();
END_IF
END_METHOD

PROPERTY StateID : STRING
GET
StateID := 'Set Ha Offset State';
END_GET
END_PROPERTY

METHOD ToIdle : BOOL
IF NOT bBlockChange THEN
	Stage := 0;
	tonDelay(IN:=FALSE);
	tonCount(IN:=FALSE);
	bToIdle := FALSE;
	pPendant^.SetState(pPendant^.fbPendantIdleState);
ELSE
	bToIdle := TRUE;
END_IF
END_METHOD

END_FUNCTION_BLOCK

// ---- POUs/PendantControl/States/FB_PendantSetFocusState.TcPOU
FUNCTION_BLOCK FB_PendantSetFocusState EXTENDS FB_PendantState
VAR_INPUT
END_VAR
VAR_OUTPUT
END_VAR
VAR
	Stage 					: UINT;
	tonCount 				: TON:= (PT:=T#1S);
	fCurrentFocusPosition 	: LREAL;
	fSmallStep				: LREAL := 0.1;
	fBigStep				: LREAL := 1.0;
	fSetFocusPosition		: LREAL;
	sSetFocusPosition		: STRING;
	nFocusRightLength 		: UINT;
	
	bBlockChange			: BOOL := FALSE;
	bToIdle					: BOOL := FALSE;
	//Hex stuff
	aTxHexData				: ARRAY[0..2] OF BYTE;
	tonDelay				: TON:= (PT:=T#20MS);
END_VAR

METHOD FoundError : BOOL
Stage := 0;
tonDelay(IN:=FALSE);
tonCount(IN:=FALSE);
pPendant^.SetState(pPendant^.fbPendantErrorState);
END_METHOD

METHOD RunState : BOOL
CASE Stage OF
	0:
		fCurrentFocusPosition := F_RoundLREAL(pPendant^.ipFocus.Position,3);
		IF pPendant^._FastMove THEN
			IF pPendant^._MovePositive THEN
				fSetFocusPosition := fCurrentFocusPosition + fBigStep;
			ELSE
				fSetFocusPosition := fCurrentFocusPosition - fBigStep;
			END_IF
		ELSE
			IF pPendant^._MovePositive THEN
				fSetFocusPosition := fCurrentFocusPosition + fSmallStep;
			ELSE
				fSetFocusPosition := fCurrentFocusPosition - fSmallStep;
			END_IF
		END_IF
		pPendant^.ipFocus.Position := fSetFocusPosition;
		Stage := Stage +1;
	1:
		// Block State Change while full text is send -> to not run into issues with commands
		// Does not include Error State
		bBlockChange := TRUE;
		IF NOT pPendant^.fbSendHex.Busy OR pPendant^.fbSendString.Busy THEN
			Stage := Stage +1;
		END_IF
	2: 
		// send sequence for two line text. For first line: fe, 01, 00, 0c, first 8 char, second 8 char
		HEXSTR_TO_DATA('fe', ADR(aTxHexData), SIZEOF(aTxHexData));
		pPendant^.fbSendHex(
				pSendData:= ADR(aTxHexData),
				Length	:= 1,
				TXbuffer:= TxBufferPendant,
				Busy=>,
				Error=> );
		IF NOT pPendant^.fbSendHex.Busy THEN
			Stage := Stage +1;
		END_IF
	3: 
		HEXSTR_TO_DATA('01', ADR(aTxHexData), SIZEOF(aTxHexData));
		pPendant^.fbSendHex(
				pSendData:= ADR(aTxHexData),
				Length	:= 1,
				TXbuffer:= TxBufferPendant,
				Busy=>,
				Error=> );
		IF NOT pPendant^.fbSendHex.Busy THEN
			Stage := Stage +1;
		END_IF
	4: 
		HEXSTR_TO_DATA('00', ADR(aTxHexData), SIZEOF(aTxHexData));
		pPendant^.fbSendHex(
				pSendData:= ADR(aTxHexData),
				Length	:= 1,
				TXbuffer:= TxBufferPendant,
				Busy=>,
				Error=> );
		IF NOT pPendant^.fbSendHex.Busy THEN
			Stage := Stage +1;
		END_IF
	5:	
		HEXSTR_TO_DATA('0c', ADR(aTxHexData), SIZEOF(aTxHexData));
		pPendant^.fbSendHex(
				pSendData:= ADR(aTxHexData),
				Length	:= 1,
				TXbuffer:= TxBufferPendant,
				Busy=>,
				Error=> );
		IF NOT pPendant^.fbSendHex.Busy THEN
			Stage := Stage +1;
		END_IF
	6:
		// send first 8 characters
		pPendant^.fbSendString(SendString:= 'Focus 1-',
					TXbuffer:= TxBufferPendant,
					Busy=>,
					Error=> );
		IF NOT pPendant^.fbSendString.Busy  THEN
			Stage := Stage +1;
		END_IF
	7: 
		tonDelay(IN:=TRUE);
		IF tonDelay.Q THEN
			tonDelay(IN:=FALSE);
			Stage:=Stage +1;
		END_IF
	8:
		// send second characters (8 max)
		pPendant^.fbSendString(SendString:= '17mm    ',
					TXbuffer:= TxBufferPendant,
					Busy=>,
					Error=> );
		IF NOT pPendant^.fbSendString.Busy  THEN
			Stage := Stage +1;
		END_IF
	9: 
		tonDelay(IN:=TRUE);
		IF tonDelay.Q THEN
			tonDelay(IN:=FALSE);
			Stage:=Stage +1;
		END_IF
	10: 
		// second line: fe, c0, 00, 0b, first 8 char, second 8 char
		HEXSTR_TO_DATA('fe', ADR(aTxHexData), SIZEOF(aTxHexData));
		pPendant^.fbSendHex(
				pSendData:= ADR(aTxHexData),
				Length	:= 1,
				TXbuffer:= TxBufferPendant,
				Busy=>,
				Error=> );
		IF NOT pPendant^.fbSendHex.Busy THEN
			Stage := Stage +1;
		END_IF
	11: 
		HEXSTR_TO_DATA('c0', ADR(aTxHexData), SIZEOF(aTxHexData));
		pPendant^.fbSendHex(
				pSendData:= ADR(aTxHexData),
				Length	:= 1,
				TXbuffer:= TxBufferPendant,
				Busy=>,
				Error=> );
		IF NOT pPendant^.fbSendHex.Busy THEN
			Stage := Stage +1;
		END_IF
	12: 
		HEXSTR_TO_DATA('00', ADR(aTxHexData), SIZEOF(aTxHexData));
		pPendant^.fbSendHex(
				pSendData:= ADR(aTxHexData),
				Length	:= 1,
				TXbuffer:= TxBufferPendant,
				Busy=>,
				Error=> );
		IF NOT pPendant^.fbSendHex.Busy THEN
			Stage := Stage +1;
		END_IF
	13:	
		HEXSTR_TO_DATA('0b', ADR(aTxHexData), SIZEOF(aTxHexData));
		pPendant^.fbSendHex(
				pSendData:= ADR(aTxHexData),
				Length	:= 1,
				TXbuffer:= TxBufferPendant,
				Busy=>,
				Error=> );
		IF NOT pPendant^.fbSendHex.Busy THEN
			Stage := Stage +1;
		END_IF
	14:
		sSetFocusPosition := CONCAT(LREAL_TO_STRING(fSetFocusPosition),'        ');
		// send first 8 characters
		pPendant^.fbSendString(SendString:= MID(sSetFocusPosition,8,1),
					TXbuffer:= TxBufferPendant,
					Busy=>,
					Error=> );
		IF NOT pPendant^.fbSendString.Busy  THEN
			Stage := Stage +1;
		END_IF
	15: 
		tonDelay(IN:=TRUE);
		IF tonDelay.Q THEN
			tonDelay(IN:=FALSE);
			Stage:=Stage +1;
		END_IF
	16:
		pPendant^.fbSendString(SendString:= 'mm      ',
					TXbuffer:= TxBufferPendant,
					Busy=>,
					Error=> );
		IF NOT pPendant^.fbSendString.Busy  THEN
			// unblock State change
			bBlockChange := FALSE;
			Stage := Stage +1;
		END_IF
	17:
		tonCount(IN:=TRUE);
		IF tonCount.Q THEN
			tonCount(IN:=FALSE);
			//restart
			Stage:=0;
		END_IF
END_CASE

IF bToIdle THEN
	THIS^.ToIdle();
END_IF
END_METHOD

PROPERTY StateID : STRING
GET
StateID := 'Set Focus State';
END_GET
END_PROPERTY

METHOD ToIdle : BOOL
IF NOT bBlockChange THEN
	Stage := 0;
	tonDelay(IN:=FALSE);
	tonCount(IN:=FALSE);
	bToIdle := FALSE;
	pPendant^.SetState(pPendant^.fbPendantIdleState);
ELSE
	bToIdle := TRUE;
END_IF
END_METHOD

END_FUNCTION_BLOCK

// ---- POUs/PendantControl/States/FB_PendantErrorState.TcPOU
FUNCTION_BLOCK FB_PendantErrorState EXTENDS FB_PendantState
VAR_INPUT
END_VAR
VAR_OUTPUT
END_VAR
VAR
END_VAR

METHOD ResetCommand : BOOL
pPendant^._Error := FALSE;
pPendant^.SetState(pPendant^.fbPendantPreInitState);
END_METHOD


METHOD RunState : BOOL
ResetCommand();
END_METHOD

PROPERTY StateID : STRING
GET
StateID := 'Error State';
END_GET
END_PROPERTY

END_FUNCTION_BLOCK

// ---- POUs/FB_SafetyHandling.TcPOU
FUNCTION_BLOCK FB_SafetyHandling
VAR
	// power on delay

	inError					AT%I*:	BOOL;		// Safety Error Condition
	outRun					AT%Q*:	BOOL;		// Run/Stop Safety
	outRestart				AT%Q*:	BOOL;		// Restart Safety
	outErrAck				AT%Q*:	BOOL;		// Error Acknowledgement 

	
	// Safety group
	fbInfoGroup1			: FB_InfoGroup;
	stInfoGroup1	AT%I*	: ST_InfoDataGroup;
	sStateGroup1			: STRING;
	
	// Estop
	fbInfoEStop1			:FB_InfoEStop;
	stInfoEStop1 	AT%I*	:ST_InfoDataFB;
	sStateEStop1			:STRING;
	sDiagEStop1				:STRING;	
	
	// Info safety inputs: unused, the EL1918's local inputs have no connection info data
	fbInfoSafetyIn			: FB_InfoConnection;
	stInfoSafetyIn 	AT%I*	: ST_InfoDataConnection;
	sStateSafetyIn			: STRING;
	sDiagSafetyIn			: STRING;
	bSafetyInCh1			: BOOL;
	bSafetyInCh2			: BOOL;
	bSafetyInCh3			: BOOL;
	bSafetyInCh4			: BOOL;
	
	// Info EL2904
	fbInfoSafetyOut			: FB_InfoConnection;
	stInfoSafetyOut AT%I*	: ST_InfoDataConnection;
	sStateSafetyOut			: STRING;
	sDiagSafetyOut			: STRING;
	bSafetyOutCh1			: BOOL;
	bSafetyOutCh2			: BOOL;
	bSafetyOutCh3			: BOOL;
	bSafetyOutCh4			: BOOL;
	
	initialStartUpStep		: INT := 0;
	startDelay 				: TON := (PT := T#2S);
	stateDelay 				: TON := (PT := T#1S);

	// #11: acknowledge on request (the telescope reset), the same ErrAck and Restart pulses as the start-up
	bAckRequest				: BOOL;			// Acknowledge() was called (one scan)
	bAckSkipped				: BOOL;			// the request was ignored this scan
	nAckStep				: INT;			// 0 idle, 1 ErrAck, 2 Restart
	ackDelay				: TON := (PT := T#1S);
	AckLog, AckSkippedLog	: FB_EventLog;

	// #59: an E-stop needs a safety acknowledge. The telescope reset fires on this flag as well as on an error,
	// so the acknowledge is not lost when the axis errors are already cleared (or never latched).
	rtrigEstop				: R_TRIG;
	bEstopDuringAck			: BOOL;			// the E-stop was pressed while an acknowledge sequence ran
	AckPendingLog			: FB_EventLog;

	
	ErrAckLog				: FB_EventLog;		// Errack logging
	RestartLog				: FB_EventLog;		// restart logging
	SafetyLog				: FB_EventLog;		// safety logging
	
	comm					: I_Comm;
END_VAR
VAR_OUTPUT
	error					: BOOL;		// error condition
	state          			: BOOL;		// safety is okay
	estop					: BOOL;		// Emergency_stop engaged
	ackPending				: BOOL;		// E-stop seen, no clean acknowledge since (#59)
	bStartUpDone			: BOOL;		// the start-up ErrAck/Restart sequence is finished (#103)
END_VAR
VAR_INPUT
	// issue a remote restart
	//remote_restart:		BOOL;
	// issue a remute run/stop
	remote_run		: BOOL := TRUE;
END_VAR

// Safety is running on start
outRun := remote_run;
GVL_Safety.Run := outRun;

// error?
error := inError;

// get safety status
fbInfoGroup1(
	stInfoData	:= stInfoGroup1,
	sState		=> sStateGroup1);
state := sStateGroup1 = 'RUN' OR initialStartUpStep <> 100;

// estop triggered?
fbInfoEStop1(
	stInfoData	:= stInfoEStop1, 
	sState		=> sStateEStop1, 
	sDiag		=> sDiagEStop1);
estop := sStateEStop1 <> 'RUN' AND initialStartUpStep = 100;

// #59: every E-stop (also one held through the PLC start, estop is masked until the start-up is done) needs an
// acknowledge. Cleared only by a clean sequence below; nothing is acknowledged automatically.
rtrigEstop(CLK := estop);
IF rtrigEstop.Q THEN
	ackPending := TRUE;
END_IF

// No info for the safety inputs: they are the EL1918's own local inputs, not an FSoE connection,
// so TwinSAFE offers no connection info data for them and stInfoSafetyIn stays unlinked (#34).

//Info SafetyOut EL2904
fbInfoSafetyOut(
	stInfoData		:=stInfoSafetyOut, 
	sState			=>sStateSafetyOut, 
	sDiag			=>sDiagSafetyOut, 
	bChannel1		=>bSafetyOutCh1, 
	bChannel2		=>bSafetyOutCh2, 
	bChannel3		=>bSafetyOutCh3, 
	bChannel4		=>bSafetyOutCh4);

// initial startup	
CASE initialStartUpStep OF
	0:
		// begin start up procedure, do ErrAck
		startDelay(IN := TRUE);
		IF startDelay.Q THEN
			startDelay(IN := FALSE);
			initialStartUpStep := initialStartUpStep+1;
		END_IF		
	1:
		// do err ack 
		GVL_Safety.ErrAck := TRUE;
		stateDelay(IN := TRUE);
		IF stateDelay.Q THEN
			stateDelay(IN := FALSE);
			GVL_Safety.ErrAck := FALSE;
			initialStartUpStep := initialStartUpStep+1;
		END_IF
	2:
		// do restart
		GVL_Safety.Restart := TRUE;
		stateDelay(IN := TRUE);
		IF stateDelay.Q THEN
			stateDelay(IN := FALSE);
			GVL_Safety.Restart := FALSE;
			initialStartUpStep := 100;
		END_IF		
END_CASE
bStartUpDone := initialStartUpStep = 100;

// #11: acknowledge on request. Ignored while the start-up runs, while a sequence runs, and while the E-stop is
// pressed (the safety logic also gates the drive acknowledge on the E-stop input, so it would do nothing).
bAckSkipped := bAckRequest AND nAckStep = 0 AND (initialStartUpStep <> 100 OR estop);
IF bAckRequest AND nAckStep = 0 AND NOT bAckSkipped THEN
	nAckStep := 1;
END_IF
bAckRequest := FALSE;

// an E-stop during the sequence spoils it: TwinSAFE gates the Restart on the E-stop input
bEstopDuringAck := bEstopDuringAck OR (estop AND nAckStep <> 0);

CASE nAckStep OF
	1:
		GVL_Safety.ErrAck := TRUE;
		ackDelay(IN := TRUE);
		IF ackDelay.Q THEN
			ackDelay(IN := FALSE);
			GVL_Safety.ErrAck := FALSE;
			nAckStep := 2;
		END_IF
	2:
		GVL_Safety.Restart := TRUE;
		ackDelay(IN := TRUE);
		IF ackDelay.Q THEN
			ackDelay(IN := FALSE);
			GVL_Safety.Restart := FALSE;
			IF NOT bEstopDuringAck THEN
				ackPending := FALSE;
			END_IF
			bEstopDuringAck := FALSE;
			nAckStep := 0;
		END_IF
END_CASE

AckLog(
	Trigger		:= nAckStep = 1,
	Level		:= ADSLOG_MSGTYPE_WARN,
	OnMessage	:= 'Safety acknowledge by telescope reset: ErrAck, then Restart.',
	Comm		:= comm);
AckSkippedLog(
	Trigger		:= bAckSkipped,
	Level		:= ADSLOG_MSGTYPE_WARN,
	OnMessage	:= 'Safety acknowledge skipped: E-stop pressed or safety start-up running.',
	Comm		:= comm);
AckPendingLog(
	Trigger		:= ackPending,
	Level		:= ADSLOG_MSGTYPE_WARN,
	OnMessage	:= 'Safety acknowledge needed after the E-stop: release it, then reset the telescope.',
	OffMessage	:= 'Safety acknowledged after the E-stop.',
	OffLevel	:= ADSLOG_MSGTYPE_HINT,
	Comm		:= comm);
(*

ErrAckLog(  
	Trigger 	:= outErrAck,
	OnMessage 	:= 'Safety error was acknowledged.',
	Comm		:= comm
);
			
RestartLog(	
	Trigger 	:= outRestart,
	Level 		:= ADSLOG_MSGTYPE_WARN,
	OnMessage 	:= 'Safety was restarted.',
	Comm		:= comm
);

SafetyLog(	
	Trigger 	:= estop,
	Level 		:= ADSLOG_MSGTYPE_ERROR,
	OnMessage 	:= 'Safety Error! Emergency stop enganged!',
	OffMessage 	:= 'Safety is OK.',
	OffLevel 	:= ADSLOG_MSGTYPE_HINT,
	Comm		:= comm);
*)

// #11: request the safety acknowledge (ErrAck 1 s, then Restart 1 s), as the telescope reset does after an E-stop
METHOD Acknowledge : BOOL
bAckRequest := TRUE;
END_METHOD

//FB_Init is always available implicitly and it is used primarily for initialization.
//The return value is not evaluated. For a specific influence, you can also declare the
//methods explicitly and provide additional code there with the standard initialization
//code. You can evaluate the return value.
METHOD FB_Init: BOOL
VAR_INPUT
    bInitRetains	: BOOL; // TRUE: the retain variables are initialized (reset warm / reset cold)
    bInCopyCode		: BOOL;  // TRUE: the instance will be copied to the copy code afterward (online change)
	comm			: I_Comm;	      
END_VAR
THIS^.comm := comm;
END_METHOD

END_FUNCTION_BLOCK

// ---- POUs/SerialBackground.TcPOU
PROGRAM SerialBackground
VAR
	fbDomeSerial : FB_SerialBackground;
	fbPendantSerial : FB_SerialBackground;
END_VAR

fbDomeSerial(RxBuffer:=RxBufferDome, TxBuffer:=TxBufferDome);

fbPendantSerial(RxBuffer:=RxBufferPendant, TxBuffer:=TxBufferPendant);

END_PROGRAM

// ---- POUs/FB_SerialBackground.TcPOU
FUNCTION_BLOCK FB_SerialBackground
VAR_IN_OUT
	TxBuffer	: ComBuffer;
	RxBuffer	: ComBuffer;
END_VAR
VAR
	(* background communication with the EL6001 terminal *)
	fbEL6001Ctrl		: SerialLineControl;
	bEL6001CtrlError	: BOOL;
	eEL6001CtrlErrorID	: ComError_t;
	(* 	I/O variables for a EL6001 terminal*)
	stIn_EL6001 AT %I*	: EL6inData22B;	(* linked to the EL6001 in the TwinCAT System Manager *)
	stOut_EL6001 AT %Q*	: EL6outData22B;(* linked to the EL6001 in the TwinCAT System Manager *)
	
	fbClear				: ClearComBuffer;
END_VAR

(*
The SerialLineControl function block is supposed to be called in every PLC cycle.
It communicates with the serial line hardware device and transmits or receives data.
The SerialLineControl can be called in the standard task (e.g.for PcCOM port usage) 
or in a separate fast task (e.g.for terminal usage) as well.
A fast separate task will be necessary at high baud rates or with KL6001 terminals 
which have a small process image (3 or 5 data bytes only)
*)

(* background communication with the EL6001 terminal *)
fbEL6001Ctrl(
	Mode:= SERIALLINEMODE_EL6_22B, 
	pComIn:= ADR(stIn_EL6001), 
	pComOut:= ADR(stOut_EL6001), 
	SizeComIn:= SIZEOF(stIn_EL6001), 
	Error=> , 
	ErrorID=> , 
	TxBuffer:= TxBuffer, 
	RxBuffer:= RxBuffer );
IF fbEL6001Ctrl.Error THEN
	bEL6001CtrlError := TRUE;
	eEL6001CtrlErrorID := fbEL6001Ctrl.ErrorID;
END_IF

fbClear(Buffer:=TxBuffer);

END_FUNCTION_BLOCK

// ---- POUs/Testing/FB_RefMarkerSearch.TcPOU
FUNCTION_BLOCK FB_RefMarkerSearch
VAR_INPUT
	Enable					: BOOL;
END_VAR
VAR_OUTPUT
END_VAR
VAR
	Axis						: AXIS_REF;
	Trigger						: TRIGGER_REF;
	bReady	: BOOL;
	btest : Bool;
	Axis_Status:	MC_ReadStatus;
	Axis_Home:		MC_Home;
	Axis_Power:		MC_Power;
	TouchProbe:		MC_TouchProbe;
	
	aRefPoints  : ARRAY [0..100] OF LREAL;
	aDistance	: ARRAY [1..100] OF LREAL;
	nIndx : UINT := 0;
	nState : UINT := 0;
	
	iErrorId					: UDINT;
	iCommandAborted				: BOOL;
END_VAR

// query the status of the axis at the beginning of the cycle
Axis_Status(Enable := TRUE,
			Axis := Axis);

// Enable the axis (power signal or manual enable)
Axis_Power(
	Axis := Axis,
	Enable := Enable,
	Enable_Positive := Enable,
	Enable_Negative := Enable,
	Override := 100.0,
	Status => bReady);

Trigger.EncoderID := 1;
Trigger.Edge := E_SignalEdge.RisingEdge;
Trigger.Mode := E_TouchProbeMode.TOUCHPROBEMODE_SINGLE_COMPATIBILITYMODE;
Trigger.TouchProbe := E_TouchProbe.TouchProbe1;
CASE nState OF
	0 :	(* init *)
		IF bReady AND btest THEN
			nIndx := 0; // reset index
			nState := nState + 1;
		END_IF
		
	1:
		TouchProbe(
			Execute 		:= TRUE,
			Axis 			:= Axis,
			TriggerInput 	:= Trigger,
			RecordedPosition => aRefPoints[nIndx]);
			
		IF NOT TouchProbe.Busy AND TouchProbe.Done THEN
			TouchProbe(	
				Execute			:= FALSE,
				TriggerInput 	:= Trigger, 
				Axis			:= Axis);
			IF nIndx > 0 THEN
				aDistance[nIndx] := F_RoundLREAL(ABS(aRefPoints[nIndx] - aRefPoints[nIndx-1]), 2);
			END_IF
			nIndx := nIndx + 1;
			nState :=  1; 	(* search for next position *)
		ELSIF NOT TouchProbe.Busy AND (TouchProbe.Error OR TouchProbe.CommandAborted) THEN
			iErrorID := TouchProbe.ErrorID;
			
			TouchProbe(	
				Execute			:= FALSE, 
				TriggerInput 	:= Trigger,
				Axis			:= Axis);

			nState 	:= 20;
		END_IF
END_CASE

END_FUNCTION_BLOCK

// ---- GlobalTextList.TcGTLO
TEXTLIST GlobalTextList
  785 = 'Azimuth:'
  815 = 'Derotator:'
  524 = 'Diag: %s'
  101 = 'EL1904'
  761 = 'EL2904'
  409 = 'Elevation:'
  868 = 'ErrAck'
  225 = 'Estop: %s'
  469 = 'Reset'
  789 = 'Restart'
  255 = 'Safety'
  521 = 'Safety Diag: %s'
  672 = 'Safety State: %s'
  809 = 'State: %s'
  328 = 'STO ErrAck:'
  488 = 'STO:'
END_TEXTLIST

// ---- VISUs/Safety.TcVIS
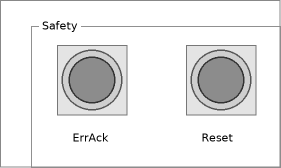
VISUALIZATION Safety  // 281x168
    GroupBox (31,18 250x150), "Safety"
        PushSwitchLed (155,27 70x70), variable: GVL_Safety.Restart, behaviour: TOGGLE, style: Switch-PushSwitchLed-Gray
        PushSwitchLed (26,27 70x70), variable: GVL_Safety.ErrAck, behaviour: TOGGLE, style: Switch-PushSwitchLed-Gray
        Label (21,105 77x30), "ErrAck"
        Label (157,105 59x30), "Reset"
END_VISUALIZATION
